      rq_wait_pos_spe_for_request(255, 204, 255, "1")
      rq_go_to("1")
      rq_wait("1")
      # end: URCap Program Node
      $ 2066 "Decap"
      $ 2067 "Action_Info≔'decapping'"
      global Action_Info="decapping"
      $ 2068 "Set GRP_3F_Enable=On"
      set_standard_digital_out(4, True)
      $ 2069 "Set GRP_3F_Decap=On"
      set_standard_digital_out(3, True)
      $ 2070 "Force"
      sleep(0.02)
      zero_ftsensor()
      force_mode(p[0.0,0.0,0.0,0.0,0.0,0.0], [0, 0, 1, 0, 0, 0], [0.0, 0.0, 1.0, 0.0, 0.0, 0.0], 2, [0.1, 0.1, 0.001, 0.3490658503988659, 0.3490658503988659, 0.3490658503988659])
      $ 2071 "check_decapping(offset=0.015, timeout=10, abort=CMD_Hold)" "noBreak"
      check_decapping(offset=0.015, timeout=10, abort=CMD_Hold)
      end_force_mode()
      stopl(5.0)
      $ 2072 "Set GRP_3F_Decap=Off"
      set_standard_digital_out(3, False)
      $ 2073 "Set GRP_3F_Enable=Off"
      set_standard_digital_out(4, False)
      $ 2074 "MoveL"
      $ 2075 "Waypoint_90" "breakAfter"
      movel(Waypoint_90_p, a=0.5, v=0.1, r=0.05)
      $ 2076 "MoveJ"
      $ 2077 "cap_dump_2" "breakAfter"
      movej(get_inverse_kin(cap_dump_2_p, qnear=cap_dump_2_q), a=0.5235987755982988, v=0.4363323129985824)
      # begin: URCap Program Node
      #   Source: Robotiq_Grippers, 3.17.0.105337, Robotiq Inc.
      #   Type: Gripper
      $ 2078 "Gripper Open (1)"
      if not(gripper_connected[0]):
        popup("Gripper 1 must be connected to run this program.", "No connection", False, True, True)
      end
      if not(rq_is_gripper_activated("1")):
        popup("Gripper 1 is not activated. Go to Installation tab > Gripper to activate it and run the program again.", "Not activated", False, True, True)
      end
      rq_set_pos_spd_for(0, 204, 255, "1")
      rq_wait_pos_spe_for_request(0, 204, 255, "1")
      rq_go_to("1")
      rq_wait("1")
      # end: URCap Program Node
      $ 2079 "MoveJ"
      $ 2080 "Waypoint_91" "breakAfter"
      movej(get_inverse_kin(Waypoint_91_p, qnear=Waypoint_91_q), a=0.5235987755982988, v=0.4363323129985824, r=0.036)
    elif (33 == switch_1):
      $ 2081 "Case 33"
      $ 2082 "Shake and liquid transfer"
      $ 2083 "MoveL"
      $ 2084 "Vial_liq_abov_1" "breakAfter"
      movel(Vial_liq_abov_1_p, a=0.5, v=0.1)
      $ 2085 "Vial_liq_pick_3" "breakAfter"
      movel(Vial_liq_pick_3_p, a=0.5, v=0.1)
      $ 2086 "Vial_liq_pick_4" "breakAfter"
      movel(Vial_liq_pick_4_p, a=0.5, v=0.1)
      # begin: URCap Program Node
      #   Source: Robotiq_Grippers, 3.17.0.105337, Robotiq Inc.
      #   Type: Gripper
      $ 2087 "Gripper Close (1)"
      if not(gripper_connected[0]):
        popup("Gripper 1 must be connected to run this program.", "No connection", False, True, True)
      end
      if not(rq_is_gripper_activated("1")):
        popup("Gripper 1 is not activated. Go to Installation tab > Gripper to activate it and run the program again.", "Not activated", False, True, True)
      end
      rq_set_pos_spd_for(255, 82, 71, "1")
      rq_wait_pos_spe_for_request(255, 82, 71, "1")
      rq_go_to("1")
      rq_wait("1")
      # end: URCap Program Node
      $ 2088 "Wait: 1.0"
      sleep(1.0)
      $ 2089 "Set GRP_3F_Open=On"
      set_standard_digital_out(5, True)
      $ 2090 "Wait: 0.5"
      sleep(0.5)
      $ 2091 "Vial_liq_abov_2" "breakAfter"
      movel(Vial_liq_abov_2_p, a=0.3, v=0.05, r=0.05)
      $ 2092 "MoveL"
      $ 2093 "Liquid_midway_1" "breakAfter"
      movel(Liquid_midway_1_p, a=0.5, v=0.1)
      $ 2094 "Loop 3 times"
      Loop_1 = 0
      while (Loop_1 < 3):
        $ 2095 "shake_3" "breakAfter"
        movel(shake_3_p, a=2.0, v=0.5)
        $ 2096 "shake_4" "breakAfter"
        movel(shake_4_p, a=2.0, v=0.5)
        Loop_1 = Loop_1 + 1
      end
      $ 2097 "drop_above_3" "breakAfter"
      movel(drop_above_3_p, a=0.5, v=0.1)
      $ 2098 "drop_above_4" "breakAfter"
      movel(drop_above_4_p, a=0.5, v=0.1)
      $ 2099 "liq_tran_3" "breakAfter"
      movel(liq_tran_3_p, a=0.5, v=0.05, r=0.008)
      $ 2100 "Wait: 1.0"
      sleep(1.0)
      $ 2101 "drop_above_5" "breakAfter"
      movel(drop_above_5_p, a=0.5, v=0.1)
      $ 2102 "Waypoint_92" "breakAfter"
      movel(Waypoint_92_p, a=0.5, v=0.1)
      $ 2103 "liq_tran_4" "breakAfter"
      movel(liq_tran_4_p, a=0.5, v=0.05)
      $ 2104 "Wait: 1.0"
      sleep(1.0)
      $ 2105 "drop_above_6" "breakAfter"
      movel(drop_above_6_p, a=0.5, v=0.1)
      $ 2106 "drop_above_7" "breakAfter"
      movel(drop_above_7_p, a=0.5, v=0.1)
      $ 2107 "Liquid_midway_2" "breakAfter"
      movel(Liquid_midway_2_p, a=0.5, v=0.1)
      $ 2108 "MoveL"
      $ 2109 "Vial_drop_abo_1" "breakAfter"
      movel(Vial_drop_abo_1_p, a=0.5, v=0.1)
      $ 2110 "Vial_liq_drop_1" "breakAfter"
      movel(Vial_liq_drop_1_p, a=0.5, v=0.1)
      # begin: URCap Program Node
      #   Source: Robotiq_Grippers, 3.17.0.105337, Robotiq Inc.
      #   Type: Gripper
      $ 2111 "Gripper Open (1)"
      if not(gripper_connected[0]):
        popup("Gripper 1 must be connected to run this program.", "No connection", False, True, True)
      end
      if not(rq_is_gripper_activated("1")):
        popup("Gripper 1 is not activated. Go to Installation tab > Gripper to activate it and run the program again.", "Not activated", False, True, True)
      end
      rq_set_pos_spd_for(0, 82, 71, "1")
      rq_wait_pos_spe_for_request(0, 82, 71, "1")
      rq_go_to("1")
      rq_wait("1")
      # end: URCap Program Node
      $ 2112 "Vial_drop_abo_2" "breakAfter"
      movel(Vial_drop_abo_2_p, a=0.5, v=0.1)
    elif (34 == switch_1):
      $ 2113 "Case 34"
      $ 2114 "Task≔'Dosing'"
      global Task="Dosing"
      $ 2115 "tilt_to_home()"
      tilt_to_home()
      $ 2116 "Powder dosing all"
      $ 2117 "tilt_angle_sent≔0.0"
      global tilt_angle_sent=0.0
      $ 2118 "send_target_info()"
      send_target_info()
      $ 2120 "prev_spat≔''"
      global prev_spat=""
      $ 2121 "spatula≔''"
      global spatula=""
      $ 2122 "scoop_status≔'normal'"
      global scoop_status="normal"
      $ 2123 "send_powder_info()"
      send_powder_info()
      $ 2124 "Set AO[0]=0.0"
      set_standard_analog_out(0, 0.0)
      $ 2125 "Wait: 0.2"
      sleep(0.2)
      $ 2126 "reach pots decapping pose"
      # begin: URCap Program Node
      #   Source: SensoPart VISOR Robotic, 2.0.6, SensoPart Industriesensorik GmbH
      #   Type: VISOR Robotic App
      $ 2132 "VISOR Easy Pick"
      def visorFuncEasyPick_e02a40():
        # begin: URCap Program Node
        #   Source: SensoPart VISOR Robotic, 2.0.6, SensoPart Industriesensorik GmbH
        #   Type: Easy Pick Setup
        $ 2133 "# 1 Setup" "noBreak"
        local easyPickVisorId = 1
        local easyPickArmMounted = True
        local easyPickSetJob = True
        local easyPickJobName = "Weight_scale"
        local easyPickAtImgAcq = False
        local easyPickImgAcqPose = Trigger
        # end: URCap Program Node
        # begin: URCap Program Node
        #   Source: SensoPart VISOR Robotic, 2.0.6, SensoPart Industriesensorik GmbH
        #   Type: Process
        $ 2134 "Process" "noBreak"
        local easyPickObjTaken = False
        local easyPickTrigger = False
        local easyPickPoseIdx = 0
        local easyPickPose = p[0,0,0,0,0,0]
        def easyPickFuncTrigger(visorId, setJob, jobName, arm):
        if (setJob):
          visor_changeJob(visorId, jobName, 6000)
        end
        if (arm):
          visor_trigger(visorId, 6000, "arm")
        else:
          visor_trigger(visorId, 6000)
        end
        global easyPickParts_4=visor_partsFound(visorId)
        visor_easyPickUpdate(visorId, "parts", visor_partsFound(visorId))
        return visor_getPose3d(visorId, 0)
      end
      while (not easyPickObjTaken):
        easyPickTrigger = (easyPickCount_4 >= visor_partsFound(easyPickVisorId)) or (easyPickCount_4 > 9) or (not visor_easyPickCheckIdent("02a34f", easyPickVisorId))
        if (easyPickTrigger):
          easyPickCount_4 = 0
        end
        easyPickPoseIdx = easyPickCount_4
        easyPickPose = visor_getPose3d(easyPickVisorId, easyPickPoseIdx)
        visor_easyPickUpdate(easyPickVisorId, "counter", easyPickPoseIdx)
        # begin: URCap Program Node
        #   Source: SensoPart VISOR Robotic, 2.0.6, SensoPart Industriesensorik GmbH
        #   Type: Image Acquisition Pose
        $ 2135 "Image Acquisition Pose" "noBreak"
        if (easyPickTrigger):
          if (not easyPickAtImgAcq):
            movej(pose_trans(easyPickImgAcqPose,p[0.0000,0.0000,-0.0000,0.0000,0.0000,0.0000]),a=1.3963,v=1.0472,t=0.000000,r=0.000000)
            easyPickAtImgAcq = True
          end
          easyPickPose = easyPickFuncTrigger(easyPickVisorId, easyPickSetJob, easyPickJobName, easyPickArmMounted)
        end
        # end: URCap Program Node
        # begin: URCap Program Node
        #   Source: SensoPart VISOR Robotic, 2.0.6, SensoPart Industriesensorik GmbH
        #   Type: Object Detected
        $ 2136 "Object Detected" "noBreak"
        if (visor_partsFound(easyPickVisorId) > 0):
          $ 2137 "Open Gripper" "noBreak"
          $ 2138 "weight_value≔get_weight()" "noBreak"
          global weight_value=get_weight()
          $ 2139 "Wait: 0.5" "noBreak"
          sleep(0.5)
          $ 2140 "diff≔target_weight-weight_value" "noBreak"
          global diff=target_weight-weight_value
          $ 2141 "compute_level_percent(W_now, weight_value)" "noBreak"
          compute_level_percent(W_now, weight_value)
          $ 2142 "send_level_info()" "noBreak"
          send_level_info()
          $ 2143 "spatula≔select_spatula(Flowability, level, diff, bulk_density, mouth_d)" "noBreak"
          global spatula=select_spatula(Flowability, level, diff, bulk_density, mouth_d)
          $ 2144 "Wait: 0.2" "noBreak"
          sleep(0.2)
          $ 2145 "send_spatula_info()" "noBreak"
          send_spatula_info()
          $ 2146 "Pick spatula" "noBreak"
          $ 2147 "If spatula ≟ 'spatula_L'" "noBreak"
          if (spatula  ==  "spatula_L"):
            $ 2148 "MoveJ" "noBreak"
            $ 2149 "Spatula_otw" "noBreak"
            movej(get_inverse_kin(Spatula_otw_p, qnear=Spatula_otw_q), a=1.3962634015954636, v=1.0471975511965976)
            $ 2150 "pick_spat_L_abv" "noBreak"
            movej(get_inverse_kin(pick_spat_L_abv_p, qnear=pick_spat_L_abv_q), a=1.3962634015954636, v=1.0471975511965976)
            $ 2151 "MoveL" "noBreak"
            $ 2152 "spat_L_pick" "noBreak"
            movel(spat_L_pick_p, a=1.2, v=0.25)
            # begin: URCap Program Node
            #   Source: Robotiq_Grippers, 3.17.0.105337, Robotiq Inc.
            #   Type: Gripper
            $ 2153 "Gripper Close (1)" "noBreak"
            if not(gripper_connected[0]):
              popup("Gripper 1 must be connected to run this program.", "No connection", False, True, True)
            end
            if not(rq_is_gripper_activated("1")):
              popup("Gripper 1 is not activated. Go to Installation tab > Gripper to activate it and run the program again.", "Not activated", False, True, True)
            end
            rq_set_pos_spd_for(255, 0, 77, "1")
            rq_wait_pos_spe_for_request(255, 0, 77, "1")
            rq_go_to("1")
            rq_wait("1")
            # end: URCap Program Node
            $ 2154 "spat_L_lift" "noBreak"
            movel(spat_L_lift_p, a=1.2, v=0.25, r=0.01)
            $ 2155 "spat_L_side" "noBreak"
            movel(spat_L_side_p, a=1.2, v=0.25, r=0.01)
            $ 2156 "spat_L_up" "noBreak"
            movel(spat_L_up_p, a=1.2, v=0.25, r=0.05)
            $ 2157 "MoveJ" "noBreak"
            $ 2158 "Spatula_otw" "noBreak"
            movej(get_inverse_kin(Spatula_otw_p, qnear=Spatula_otw_q), a=1.3962634015954636, v=1.0471975511965976)
          else:
            $ 2159 "ElseIf spatula ≟'spatula_M'" "noBreak"
            if (spatula  == "spatula_M"):
              $ 2160 "MoveJ" "noBreak"
              $ 2161 "Spatula_otw" "noBreak"
              movej(get_inverse_kin(Spatula_otw_p, qnear=Spatula_otw_q), a=1.3962634015954636, v=1.0471975511965976)
              $ 2162 "spat_M_up" "noBreak"
              movej(get_inverse_kin(spat_M_up_p, qnear=spat_M_up_q), a=1.3962634015954636, v=1.0471975511965976, r=0.05)
              $ 2163 "MoveL" "noBreak"
              $ 2164 "spat_M_pick" "noBreak"
              movel(spat_M_pick_p, a=1.2, v=0.25)
              # begin: URCap Program Node
              #   Source: Robotiq_Grippers, 3.17.0.105337, Robotiq Inc.
              #   Type: Gripper
              $ 2165 "Gripper Close (1)" "noBreak"
              if not(gripper_connected[0]):
                popup("Gripper 1 must be connected to run this program.", "No connection", False, True, True)
              end
              if not(rq_is_gripper_activated("1")):
                popup("Gripper 1 is not activated. Go to Installation tab > Gripper to activate it and run the program again.", "Not activated", False, True, True)
              end
              rq_set_pos_spd_for(255, 0, 77, "1")
              rq_wait_pos_spe_for_request(255, 0, 77, "1")
              rq_go_to("1")
              rq_wait("1")
              # end: URCap Program Node
              $ 2166 "spat_M_up" "noBreak"
              movel(spat_M_up_p, a=1.2, v=0.25, r=0.05)
              $ 2167 "Spatula_otw" "noBreak"
              movel(Spatula_otw_p, a=1.2, v=0.25)
              $ 2168 "switch_spat_M≔ False " "noBreak"
              global switch_spat_M=  False
            else:
              $ 2169 "ElseIf spatula≟'spatula_S'" "noBreak"
              if (spatula == "spatula_S"):
                $ 2170 "MoveJ" "noBreak"
                $ 2171 "Spatula_otw" "noBreak"
                movej(get_inverse_kin(Spatula_otw_p, qnear=Spatula_otw_q), a=1.3962634015954636, v=1.0471975511965976)
                $ 2172 "spat_S_Up_7" "noBreak"
                movej(get_inverse_kin(spat_S_Up_7_p, qnear=spat_S_Up_7_q), a=1.3962634015954636, v=1.0471975511965976, r=0.05)
                $ 2173 "MoveL" "noBreak"
                $ 2174 "spat_S_Pick_4" "noBreak"
                movel(spat_S_Pick_4_p, a=1.2, v=0.25)
                # begin: URCap Program Node
                #   Source: Robotiq_Grippers, 3.17.0.105337, Robotiq Inc.
                #   Type: Gripper
                $ 2175 "Gripper Close (1)" "noBreak"
                if not(gripper_connected[0]):
                  popup("Gripper 1 must be connected to run this program.", "No connection", False, True, True)
                end
                if not(rq_is_gripper_activated("1")):
                  popup("Gripper 1 is not activated. Go to Installation tab > Gripper to activate it and run the program again.", "Not activated", False, True, True)
                end
                rq_set_pos_spd_for(255, 0, 77, "1")
                rq_wait_pos_spe_for_request(255, 0, 77, "1")
                rq_go_to("1")
                rq_wait("1")
                # end: URCap Program Node
                $ 2176 "spat_S_Up_8" "noBreak"
                movel(spat_S_Up_8_p, a=1.2, v=0.25, r=0.05)
                $ 2177 "Spatula_otw" "noBreak"
                movel(Spatula_otw_p, a=1.2, v=0.25)
                $ 2178 "switch_spat_S≔ False " "noBreak"
                global switch_spat_S=  False
              else:
                $ 2179 "ElseIf spatula≟'spatula_flat_M'" "noBreak"
                if (spatula == "spatula_flat_M"):
                  $ 2180 "MoveJ" "noBreak"
                  $ 2181 "Spatula_otw" "noBreak"
                  movej(get_inverse_kin(Spatula_otw_p, qnear=Spatula_otw_q), a=1.3962634015954636, v=1.0471975511965976)
                  $ 2182 "spat_flatM_up" "noBreak"
                  movej(get_inverse_kin(spat_flatM_up_p, qnear=spat_flatM_up_q), a=1.3962634015954636, v=1.0471975511965976, r=0.05)
                  $ 2183 "MoveL" "noBreak"
                  $ 2184 "spat_flatM_pick" "noBreak"
                  movel(spat_flatM_pick_p, a=1.2, v=0.25)
                  # begin: URCap Program Node
                  #   Source: Robotiq_Grippers, 3.17.0.105337, Robotiq Inc.
                  #   Type: Gripper
                  $ 2185 "Gripper Close (1)" "noBreak"
                  if not(gripper_connected[0]):
                    popup("Gripper 1 must be connected to run this program.", "No connection", False, True, True)
                  end
                  if not(rq_is_gripper_activated("1")):
                    popup("Gripper 1 is not activated. Go to Installation tab > Gripper to activate it and run the program again.", "Not activated", False, True, True)
                  end
                  rq_set_pos_spd_for(255, 0, 77, "1")
                  rq_wait_pos_spe_for_request(255, 0, 77, "1")
                  rq_go_to("1")
                  rq_wait("1")
                  # end: URCap Program Node
                  $ 2186 "spat_flatM_up" "noBreak"
                  movel(spat_flatM_up_p, a=1.2, v=0.25, r=0.05)
                  $ 2187 "Spatula_otw" "noBreak"
                  movel(Spatula_otw_p, a=1.2, v=0.25)
                  $ 2188 "switch_spat_F_M≔ False " "noBreak"
                  global switch_spat_F_M=  False
                else:
                  $ 2189 "ElseIf spatula≟'spatula_flat_S'" "noBreak"
                  if (spatula == "spatula_flat_S"):
                    $ 2190 "MoveJ" "noBreak"
                    $ 2191 "Spatula_otw" "noBreak"
                    movej(get_inverse_kin(Spatula_otw_p, qnear=Spatula_otw_q), a=1.3962634015954636, v=1.0471975511965976)
                    $ 2192 "spat_flatS_up" "noBreak"
                    movej(get_inverse_kin(spat_flatS_up_p, qnear=spat_flatS_up_q), a=1.3962634015954636, v=1.0471975511965976, r=0.05)
                    $ 2193 "MoveL" "noBreak"
                    $ 2194 "spat_flatS_pick" "noBreak"
                    movel(spat_flatS_pick_p, a=1.2, v=0.25)
                    # begin: URCap Program Node
                    #   Source: Robotiq_Grippers, 3.17.0.105337, Robotiq Inc.
                    #   Type: Gripper
                    $ 2195 "Gripper Close (1)" "noBreak"
                    if not(gripper_connected[0]):
                      popup("Gripper 1 must be connected to run this program.", "No connection", False, True, True)
                    end
                    if not(rq_is_gripper_activated("1")):
                      popup("Gripper 1 is not activated. Go to Installation tab > Gripper to activate it and run the program again.", "Not activated", False, True, True)
                    end
                    rq_set_pos_spd_for(255, 0, 77, "1")
                    rq_wait_pos_spe_for_request(255, 0, 77, "1")
                    rq_go_to("1")
                    rq_wait("1")
                    # end: URCap Program Node
                    $ 2196 "spat_flatS_up" "noBreak"
                    movel(spat_flatS_up_p, a=1.2, v=0.25, r=0.05)
                    $ 2197 "Spatula_otw" "noBreak"
                    movel(Spatula_otw_p, a=1.2, v=0.25)
                    $ 2198 "switch_spat_F_S≔ False " "noBreak"
                    global switch_spat_F_S=  False
                  end
                end
              end
            end
          end
          $ 2199 "Action_Info≔'Scooping'" "noBreak"
          global Action_Info="Scooping"
          $ 2200 "auto_tilt_and_scoop(W_now, target_weight, weight_value)" "noBreak"
          auto_tilt_and_scoop(W_now, target_weight, weight_value)
          $ 2201 "Action_Info≔'Dosing'" "noBreak"
          global Action_Info="Dosing"
          # begin: URCap Program Node
          #   Source: SensoPart VISOR Robotic, 2.0.6, SensoPart Industriesensorik GmbH
          #   Type: Approach Pose
          $ 2202 "Approach Pose" "noBreak"
          movej(pose_trans(easyPickPose,p[0.0000,0.0000,-0.0000,0.0000,0.0000,0.0000]),a=0.2618,v=0.1745,t=0.000000,r=0.000000)
          # end: URCap Program Node
          # begin: URCap Program Node
          #   Source: SensoPart VISOR Robotic, 2.0.6, SensoPart Industriesensorik GmbH
          #   Type: Target Pose
          $ 2203 "Target Pose" "noBreak"
          movel(pose_trans(easyPickPose,p[0.0000,0.0000,-0.0000,0.0000,0.0000,0.0000]),a=0.0500,v=0.0200,t=0.000000,r=0.000000)
          # end: URCap Program Node
          $ 2204 "Close Gripper" "noBreak"
          $ 2205 "current_p≔get_actual_tcp_pose()" "noBreak"
          global current_p= get_actual_tcp_pose ()
          $ 2206 "dispense_pos≔pose_trans(current_p,p[0,0,0,0,-deg2rad(spatula_ry),0])" "noBreak"
          global dispense_pos=pose_trans(current_p,p[0,0,0,0,-deg2rad(spatula_ry),0])
          $ 2207 "Loop weight_value≤target_weight and delta_count≤3" "noBreak"
          thread Thread_while_2207():
            while (True):
              $ 2208 "MoveL" "noBreak"
              $ 2209 "dispense_pos" "noBreak"
              movel(dispense_pos, a=0.2, v=0.1)
              $ 2210 "log_weight()" "noBreak"
              log_weight()
              $ 2212 "CCW_full_Rotate()" "noBreak"
              CCW_full_Rotate()
              $ 2213 "Start_thread≔ True " "noBreak"
              global Start_thread=  True
              $ 2214 "vib_thread≔ True " "noBreak"
              global vib_thread=  True
              $ 2215 "Wait: 0.5" "noBreak"
              sleep(0.5)
              $ 2216 "If diff ≥(target_g*1.2)" "noBreak"
              if (diff  >= (target_g*1.2)):
                $ 2217 "tilt_pose≔pose_trans(get_actual_tcp_pose(), p[0, 0, 0, 0, 0, 2.0])" "noBreak"
                global tilt_pose=pose_trans(get_actual_tcp_pose(), p[0, 0, 0, 0, 0, 2.0])
                $ 2218 "movel(tilt_pose, a=0.5, v=0.5, r=0.00001)" "noBreak"
                movel(tilt_pose, a=0.5, v=0.5, r=0.00001)
              else:
                $ 2219 "Else" "noBreak"
                $ 2220 "Loop weight_value≤(target_weight-0.00) and tilt_angle≥(-1.999) and tilt_angle≤0.5" "noBreak"
                thread Thread_while_2220():
                  while (True):
                    $ 2221 "current_error≔target_weight-weight_value" "noBreak"
                    global current_error=target_weight-weight_value
                    $ 2222 "Integral_error≔Integral_error+current_error*dt" "noBreak"
                    global Integral_error=Integral_error+current_error*dt
                    $ 2223 "derivative≔(current_error-previous_error)/dt" "noBreak"
                    global derivative=(current_error-previous_error)/dt
                    $ 2224 "tilt_increment≔(kp*current_error)+(ki*Integral_error)+(kd*derivative)" "noBreak"
                    global tilt_increment=(kp*current_error)+(ki*Integral_error)+(kd*derivative)
                    $ 2225 "current_pose≔get_actual_tcp_pose()" "noBreak"
                    global current_pose= get_actual_tcp_pose ()
                    $ 2226 "tilt_angle≔current_pose[5]" "noBreak"
                    global tilt_angle=current_pose[5]
                    $ 2227 "tilt_pose≔pose_trans(current_pose, p[0, 0, 0, 0, 0, tilt_increment])" "noBreak"
                    global tilt_pose=pose_trans(current_pose, p[0, 0, 0, 0, 0, tilt_increment])
                    $ 2228 "movel(tilt_pose, a=0.1, v=0.1, r=0.00001)" "noBreak"
                    movel(tilt_pose, a=0.1, v=0.1, r=0.00001)
                    $ 2229 "previous_error≔current_error" "noBreak"
                    global previous_error=current_error
                  end
                end
                if (weight_value <= (target_weight-0.00)  and  tilt_angle >= (-1.999)  and  tilt_angle <= 0.5):
                  global thread_handler_2220=run Thread_while_2220()
                  while (weight_value <= (target_weight-0.00)  and  tilt_angle >= (-1.999)  and  tilt_angle <= 0.5):
                    sync()
                  end
                  kill thread_handler_2220
                end
              end
              $ 2230 "weight_value≔get_weight()" "noBreak"
              global weight_value=get_weight()
              $ 2231 "tilt_angle≔-1" "noBreak"
              global tilt_angle=-1
              $ 2232 "Wait: 0.5" "noBreak"
              sleep(0.5)
              $ 2233 "Start_thread≔ False " "noBreak"
              global Start_thread=  False
              $ 2234 "vib_thread≔ False " "noBreak"
              global vib_thread=  False
              $ 2235 "dispense_pos" "noBreak"
              movel(dispense_pos, a=1.2, v=0.25)
              $ 2236 "compute_level_percent(W_now, weight_value)" "noBreak"
              compute_level_percent(W_now, weight_value)
              $ 2237 "If delta<0.01" "noBreak"
              if (delta<0.01):
                $ 2238 "delta_count≔delta_count+1" "noBreak"
                global delta_count=delta_count+1
              else:
                $ 2239 "Else" "noBreak"
                $ 2240 "delta_count≔0" "noBreak"
                global delta_count=0
              end
              $ 2241 "prev_spat≔spatula" "noBreak"
              global prev_spat=spatula
              $ 2242 "Wait: 0.2" "noBreak"
              sleep(0.2)
              $ 2243 "spatula≔select_spatula(Flowability, level, diff, bulk_density, mouth_d)" "noBreak"
              global spatula=select_spatula(Flowability, level, diff, bulk_density, mouth_d)
              $ 2244 "Wait: 1.0" "noBreak"
              sleep(1.0)
              $ 2245 "send_level_info()" "noBreak"
              send_level_info()
              $ 2246 "send_spatula_info()" "noBreak"
              send_spatula_info()
              $ 2247 "Integral_error≔0" "noBreak"
              global Integral_error=0
              $ 2248 "current_error≔0" "noBreak"
              global current_error=0
              $ 2249 "previous_error≔0" "noBreak"
              global previous_error=0
              $ 2250 "Set AO[0]=0.0" "noBreak"
              set_standard_analog_out(0, 0.0)
              $ 2251 "Wait: 0.5" "noBreak"
              sleep(0.5)
              $ 2252 "swtich spatula" "noBreak"
              $ 2253 "If spatula ≟ 'spatula_M' and switch_spat_M≟ True " "noBreak"
              if (spatula  ==  "spatula_M"  and  switch_spat_M ==   True  ):
                $ 2254 "MoveJ" "noBreak"
                $ 2255 "Spatula_otw" "noBreak"
                movej(get_inverse_kin(Spatula_otw_p, qnear=Spatula_otw_q), a=1.3962634015954636, v=1.0471975511965976)
                $ 2256 "spat_L_up" "noBreak"
                movej(get_inverse_kin(spat_L_up_p, qnear=spat_L_up_q), a=1.3962634015954636, v=1.0471975511965976)
                $ 2257 "MoveL" "noBreak"
                $ 2258 "spat_L_side" "noBreak"
                movel(spat_L_side_p, a=1.2, v=0.25)
                $ 2259 "spat_L_lift" "noBreak"
                movel(spat_L_lift_p, a=1.2, v=0.25)
                $ 2260 "spat_L_pick" "noBreak"
                movel(spat_L_pick_p, a=0.2, v=0.1)
                # begin: URCap Program Node
                #   Source: Robotiq_Grippers, 3.17.0.105337, Robotiq Inc.
                #   Type: Gripper
                $ 2261 "Gripper Open (1)" "noBreak"
                if not(gripper_connected[0]):
                  popup("Gripper 1 must be connected to run this program.", "No connection", False, True, True)
                end
                if not(rq_is_gripper_activated("1")):
                  popup("Gripper 1 is not activated. Go to Installation tab > Gripper to activate it and run the program again.", "Not activated", False, True, True)
                end
                rq_set_pos_spd_for(0, 255, 77, "1")
                rq_wait_pos_spe_for_request(0, 255, 77, "1")
                rq_go_to("1")
                rq_wait("1")
                # end: URCap Program Node
                $ 2262 "spat_M_pick" "noBreak"
                movel(spat_M_pick_p, a=1.2, v=0.25)
                # begin: URCap Program Node
                #   Source: Robotiq_Grippers, 3.17.0.105337, Robotiq Inc.
                #   Type: Gripper
                $ 2263 "Gripper Close (1)" "noBreak"
                if not(gripper_connected[0]):
                  popup("Gripper 1 must be connected to run this program.", "No connection", False, True, True)
                end
                if not(rq_is_gripper_activated("1")):
                  popup("Gripper 1 is not activated. Go to Installation tab > Gripper to activate it and run the program again.", "Not activated", False, True, True)
                end
                rq_set_pos_spd_for(255, 0, 77, "1")
                rq_wait_pos_spe_for_request(255, 0, 77, "1")
                rq_go_to("1")
                rq_wait("1")
                # end: URCap Program Node
                $ 2264 "spat_M_up" "noBreak"
                movel(spat_M_up_p, a=1.2, v=0.25)
                $ 2265 "Spatula_otw" "noBreak"
                movel(Spatula_otw_p, a=1.2, v=0.25)
                $ 2266 "switch_spat_M≔ False " "noBreak"
                global switch_spat_M=  False
                $ 2267 "correction_reset()" "noBreak"
                correction_reset()
              else:
                $ 2268 "ElseIf spatula ≟ 'spatula_S' and switch_spat_S ≟ True and prev_spat≟'spatula_M'" "noBreak"
                if (spatula  ==  "spatula_S" and switch_spat_S  ==   True  and prev_spat == "spatula_M"):
                  $ 2269 "MoveL" "noBreak"
                  $ 2270 "Spatula_otw" "noBreak"
                  movel(Spatula_otw_p, a=1.2, v=0.25)
                  $ 2271 "spat_M_up" "noBreak"
                  movel(spat_M_up_p, a=1.2, v=0.25)
                  $ 2272 "spat_M_pick" "noBreak"
                  movel(spat_M_pick_p, a=0.2, v=0.1)
                  # begin: URCap Program Node
                  #   Source: Robotiq_Grippers, 3.17.0.105337, Robotiq Inc.
                  #   Type: Gripper
                  $ 2273 "Gripper Open (1)" "noBreak"
                  if not(gripper_connected[0]):
                    popup("Gripper 1 must be connected to run this program.", "No connection", False, True, True)
                  end
                  if not(rq_is_gripper_activated("1")):
                    popup("Gripper 1 is not activated. Go to Installation tab > Gripper to activate it and run the program again.", "Not activated", False, True, True)
                  end
                  rq_set_pos_spd_for(0, 255, 77, "1")
                  rq_wait_pos_spe_for_request(0, 255, 77, "1")
                  rq_go_to("1")
                  rq_wait("1")
                  # end: URCap Program Node
                  $ 2274 "spat_S_pick" "noBreak"
                  movel(spat_S_pick_p, a=1.2, v=0.25)
                  # begin: URCap Program Node
                  #   Source: Robotiq_Grippers, 3.17.0.105337, Robotiq Inc.
                  #   Type: Gripper
                  $ 2275 "Gripper Close (1)" "noBreak"
                  if not(gripper_connected[0]):
                    popup("Gripper 1 must be connected to run this program.", "No connection", False, True, True)
                  end
                  if not(rq_is_gripper_activated("1")):
                    popup("Gripper 1 is not activated. Go to Installation tab > Gripper to activate it and run the program again.", "Not activated", False, True, True)
                  end
                  rq_set_pos_spd_for(255, 0, 77, "1")
                  rq_wait_pos_spe_for_request(255, 0, 77, "1")
                  rq_go_to("1")
                  rq_wait("1")
                  # end: URCap Program Node
                  $ 2276 "spat_S_up" "noBreak"
                  movel(spat_S_up_p, a=1.2, v=0.25)
                  $ 2277 "Spatula_otw" "noBreak"
                  movel(Spatula_otw_p, a=1.2, v=0.25)
                  $ 2278 "switch_spat_S≔ False " "noBreak"
                  global switch_spat_S=  False
                  $ 2279 "correction_reset()" "noBreak"
                  correction_reset()
                else:
                  $ 2280 "ElseIf spatula≟'spatula_S' and switch_spat_S≟ True  and prev_spat≟'spatula_L'" "noBreak"
                  if (spatula == "spatula_S" and switch_spat_S ==   True    and  prev_spat == "spatula_L"):
                    $ 2281 "MoveJ" "noBreak"
                    $ 2282 "Spatula_otw" "noBreak"
                    movej(get_inverse_kin(Spatula_otw_p, qnear=Spatula_otw_q), a=1.3962634015954636, v=1.0471975511965976)
                    $ 2283 "spat_L_up" "noBreak"
                    movej(get_inverse_kin(spat_L_up_p, qnear=spat_L_up_q), a=1.3962634015954636, v=1.0471975511965976)
                    $ 2284 "MoveL" "noBreak"
                    $ 2285 "spat_L_side" "noBreak"
                    movel(spat_L_side_p, a=1.2, v=0.25)
                    $ 2286 "spat_L_lift" "noBreak"
                    movel(spat_L_lift_p, a=1.2, v=0.25)
                    $ 2287 "spat_L_pick" "noBreak"
                    movel(spat_L_pick_p, a=0.2, v=0.1)
                    # begin: URCap Program Node
                    #   Source: Robotiq_Grippers, 3.17.0.105337, Robotiq Inc.
                    #   Type: Gripper
                    $ 2288 "Gripper Open (1)" "noBreak"
                    if not(gripper_connected[0]):
                      popup("Gripper 1 must be connected to run this program.", "No connection", False, True, True)
                    end
                    if not(rq_is_gripper_activated("1")):
                      popup("Gripper 1 is not activated. Go to Installation tab > Gripper to activate it and run the program again.", "Not activated", False, True, True)
                    end
                    rq_set_pos_spd_for(0, 255, 77, "1")
                    rq_wait_pos_spe_for_request(0, 255, 77, "1")
                    rq_go_to("1")
                    rq_wait("1")
                    # end: URCap Program Node
                    $ 2289 "spat_S_pick" "noBreak"
                    movel(spat_S_pick_p, a=1.2, v=0.25)
                    # begin: URCap Program Node
                    #   Source: Robotiq_Grippers, 3.17.0.105337, Robotiq Inc.
                    #   Type: Gripper
                    $ 2290 "Gripper Close (1)" "noBreak"
                    if not(gripper_connected[0]):
                      popup("Gripper 1 must be connected to run this program.", "No connection", False, True, True)
                    end
                    if not(rq_is_gripper_activated("1")):
                      popup("Gripper 1 is not activated. Go to Installation tab > Gripper to activate it and run the program again.", "Not activated", False, True, True)
                    end
                    rq_set_pos_spd_for(255, 0, 77, "1")
                    rq_wait_pos_spe_for_request(255, 0, 77, "1")
                    rq_go_to("1")
                    rq_wait("1")
                    # end: URCap Program Node
                    $ 2291 "spat_S_up" "noBreak"
                    movel(spat_S_up_p, a=1.2, v=0.25)
                    $ 2292 "Spatula_otw" "noBreak"
                    movel(Spatula_otw_p, a=1.2, v=0.25)
                    $ 2293 "switch_spat_S≔ False " "noBreak"
                    global switch_spat_S=  False
                    $ 2294 "correction_reset()" "noBreak"
                    correction_reset()
                  else:
                    $ 2295 "ElseIf spatula≟'spatula_flat_S'  and switch_spat_F_S ≟ True " "noBreak"
                    if (spatula == "spatula_flat_S"   and  switch_spat_F_S  ==   True  ):
                      $ 2296 "MoveL" "noBreak"
                      $ 2297 "Spatula_otw" "noBreak"
                      movel(Spatula_otw_p, a=1.2, v=0.25)
                      $ 2298 "spat_flatM_up" "noBreak"
                      movel(spat_flatM_up_p, a=1.2, v=0.25)
                      $ 2299 "spat_flatM_pick" "noBreak"
                      movel(spat_flatM_pick_p, a=0.2, v=0.1)
                      # begin: URCap Program Node
                      #   Source: Robotiq_Grippers, 3.17.0.105337, Robotiq Inc.
                      #   Type: Gripper
                      $ 2300 "Gripper Open (1)" "noBreak"
                      if not(gripper_connected[0]):
                        popup("Gripper 1 must be connected to run this program.", "No connection", False, True, True)
                      end
                      if not(rq_is_gripper_activated("1")):
                        popup("Gripper 1 is not activated. Go to Installation tab > Gripper to activate it and run the program again.", "Not activated", False, True, True)
                      end
                      rq_set_pos_spd_for(0, 255, 74, "1")
                      rq_wait_pos_spe_for_request(0, 255, 74, "1")
                      rq_go_to("1")
                      rq_wait("1")
                      # end: URCap Program Node
                      $ 2301 "spat_flatS_pick" "noBreak"
                      movel(spat_flatS_pick_p, a=1.2, v=0.25)
                      # begin: URCap Program Node
                      #   Source: Robotiq_Grippers, 3.17.0.105337, Robotiq Inc.
                      #   Type: Gripper
                      $ 2302 "Gripper Close (1)" "noBreak"
                      if not(gripper_connected[0]):
                        popup("Gripper 1 must be connected to run this program.", "No connection", False, True, True)
                      end
                      if not(rq_is_gripper_activated("1")):
                        popup("Gripper 1 is not activated. Go to Installation tab > Gripper to activate it and run the program again.", "Not activated", False, True, True)
                      end
                      rq_set_pos_spd_for(255, 0, 77, "1")
                      rq_wait_pos_spe_for_request(255, 0, 77, "1")
                      rq_go_to("1")
                      rq_wait("1")
                      # end: URCap Program Node
                      $ 2303 "spat_flatS_up" "noBreak"
                      movel(spat_flatS_up_p, a=1.2, v=0.25)
                      $ 2304 "Spatula_otw" "noBreak"
                      movel(Spatula_otw_p, a=1.2, v=0.25)
                      $ 2305 "switch_spat_F_S≔ False " "noBreak"
                      global switch_spat_F_S=  False
                      $ 2306 "correction_reset()" "noBreak"
                      correction_reset()
                    end
                  end
                end
              end
              $ 2307 "tilt(level)" "noBreak"
              tilt(level)
              $ 2308 "Action_Info≔'Scooping'" "noBreak"
              global Action_Info="Scooping"
              $ 2309 "auto_tilt_and_scoop(W_now, target_weight, weight_value)" "noBreak"
              auto_tilt_and_scoop(W_now, target_weight, weight_value)
              $ 2310 "Action_Info≔'Dosing'" "noBreak"
              global Action_Info="Dosing"
            end
          end
          if (weight_value <= target_weight and delta_count <= 3):
            global thread_handler_2207=run Thread_while_2207()
            while (weight_value <= target_weight and delta_count <= 3):
              sync()
            end
            kill thread_handler_2207
          end
          $ 2311 "Start_thread≔ False " "noBreak"
          global Start_thread=  False
          $ 2312 "vib_thread≔ False " "noBreak"
          global vib_thread=  False
          # begin: URCap Program Node
          #   Source: SensoPart VISOR Robotic, 2.0.6, SensoPart Industriesensorik GmbH
          #   Type: Exit Pose
          $ 2313 "Exit Pose" "noBreak"
          movel(pose_trans(easyPickPose,p[0.0000,0.0000,-0.0000,0.0000,0.0000,0.0000]),a=0.5000,v=0.2500,t=0.000000,r=0.000000)
          # end: URCap Program Node
          easyPickObjTaken = True
        end
        # end: URCap Program Node
        # begin: URCap Program Node
        #   Source: SensoPart VISOR Robotic, 2.0.6, SensoPart Industriesensorik GmbH
        #   Type: No Object Detected
        $ 2314 "No Object Detected" "noBreak"
        if (visor_partsFound(easyPickVisorId) < 1):
          $ 2315 "Popup: No weigh scale detected" "noBreak"
          popup("No weigh scale detected", "Message", False, False, blocking=True)
          else:
        end
        # end: URCap Program Node
      end
      easyPickCount_4 = easyPickCount_4 + 1
      visor_easyPickUpdate(easyPickVisorId, "counter", easyPickCount_4)
      visor_easyPickSetIdent("02a34f", easyPickVisorId)
      # end: URCap Program Node
    end
    visorFuncEasyPick_e02a40()
    # end: URCap Program Node
    $ 2316 "MoveL"
    $ 2317 "dispense_pos" "breakAfter"
    movel(dispense_pos, a=0.2, v=0.1)
    $ 2318 "after_scoop()"
    after_scoop()
    $ 2319 "Place spatula back to the rack"
    $ 2320 "If spatula ≟ 'spatula_L'"
    if (spatula  ==  "spatula_L"):
      $ 2321 "MoveJ"
      $ 2322 "Spatula_otw" "breakAfter"
      movej(get_inverse_kin(Spatula_otw_p, qnear=Spatula_otw_q), a=1.3962634015954636, v=1.0471975511965976)
      $ 2323 "MoveL"
      $ 2324 "spat_L_up" "breakAfter"
      movel(spat_L_up_p, a=1.2, v=0.25, r=0.05)
      $ 2325 "spat_L_side" "breakAfter"
      movel(spat_L_side_p, a=1.2, v=0.25, r=0.01)
      $ 2326 "spat_L_lift" "breakAfter"
      movel(spat_L_lift_p, a=1.2, v=0.25, r=0.01)
      $ 2327 "spat_L_pick" "breakAfter"
      movel(spat_L_pick_p, a=0.2, v=0.1)
      # begin: URCap Program Node
      #   Source: Robotiq_Grippers, 3.17.0.105337, Robotiq Inc.
      #   Type: Gripper
      $ 2328 "Gripper Open (1)"
      if not(gripper_connected[0]):
        popup("Gripper 1 must be connected to run this program.", "No connection", False, True, True)
      end
      if not(rq_is_gripper_activated("1")):
        popup("Gripper 1 is not activated. Go to Installation tab > Gripper to activate it and run the program again.", "Not activated", False, True, True)
      end
      rq_set_pos_spd_for(0, 128, 128, "1")
      rq_wait_pos_spe_for_request(0, 128, 128, "1")
      rq_go_to("1")
      rq_wait("1")
      # end: URCap Program Node
      $ 2329 "MoveJ"
      $ 2330 "pick_spat_L_abv" "breakAfter"
      movej(get_inverse_kin(pick_spat_L_abv_p, qnear=pick_spat_L_abv_q), a=1.3962634015954636, v=1.0471975511965976)
      $ 2331 "Spatula_otw" "breakAfter"
      movej(get_inverse_kin(Spatula_otw_p, qnear=Spatula_otw_q), a=1.3962634015954636, v=1.0471975511965976)
    else:
      $ 2332 "ElseIf spatula ≟'spatula_M'"
      if (spatula  == "spatula_M"):
        $ 2333 "MoveJ"
        $ 2334 "Spatula_otw" "breakAfter"
        movej(get_inverse_kin(Spatula_otw_p, qnear=Spatula_otw_q), a=1.3962634015954636, v=1.0471975511965976)
        $ 2335 "spat_M_up" "breakAfter"
        movej(get_inverse_kin(spat_M_up_p, qnear=spat_M_up_q), a=1.3962634015954636, v=1.0471975511965976, r=0.05)
        $ 2336 "MoveL"
        $ 2337 "spat_M_pick" "breakAfter"
        movel(spat_M_pick_p, a=0.2, v=0.1)
        # begin: URCap Program Node
        #   Source: Robotiq_Grippers, 3.17.0.105337, Robotiq Inc.
        #   Type: Gripper
        $ 2338 "Gripper Open (1)"
        if not(gripper_connected[0]):
          popup("Gripper 1 must be connected to run this program.", "No connection", False, True, True)
        end
        if not(rq_is_gripper_activated("1")):
          popup("Gripper 1 is not activated. Go to Installation tab > Gripper to activate it and run the program again.", "Not activated", False, True, True)
        end
        rq_set_pos_spd_for(0, 128, 128, "1")
        rq_wait_pos_spe_for_request(0, 128, 128, "1")
        rq_go_to("1")
        rq_wait("1")
        # end: URCap Program Node
        $ 2339 "spat_M_up" "breakAfter"
        movel(spat_M_up_p, a=1.2, v=0.25, r=0.05)
        $ 2340 "Spatula_otw" "breakAfter"
        movel(Spatula_otw_p, a=1.2, v=0.25)
        $ 2341 "switch_spat_M≔ False "
        global switch_spat_M=  False
      else:
        $ 2342 "ElseIf spatula≟'spatula_S'"
        if (spatula == "spatula_S"):
          $ 2343 "MoveJ"
          $ 2344 "Spatula_otw" "breakAfter"
          movej(get_inverse_kin(Spatula_otw_p, qnear=Spatula_otw_q), a=1.3962634015954636, v=1.0471975511965976)
          $ 2345 "spat_S_Up_7" "breakAfter"
          movej(get_inverse_kin(spat_S_Up_7_p, qnear=spat_S_Up_7_q), a=1.3962634015954636, v=1.0471975511965976, r=0.05)
          $ 2346 "MoveL"
          $ 2347 "spat_S_Pick_4" "breakAfter"
          movel(spat_S_Pick_4_p, a=0.2, v=0.1)
          # begin: URCap Program Node
          #   Source: Robotiq_Grippers, 3.17.0.105337, Robotiq Inc.
          #   Type: Gripper
          $ 2348 "Gripper Open (1)"
          if not(gripper_connected[0]):
            popup("Gripper 1 must be connected to run this program.", "No connection", False, True, True)
          end
          if not(rq_is_gripper_activated("1")):
            popup("Gripper 1 is not activated. Go to Installation tab > Gripper to activate it and run the program again.", "Not activated", False, True, True)
          end
          rq_set_pos_spd_for(0, 255, 51, "1")
          rq_wait_pos_spe_for_request(0, 255, 51, "1")
          rq_go_to("1")
          rq_wait("1")
          # end: URCap Program Node
          $ 2349 "spat_S_Up_8" "breakAfter"
          movel(spat_S_Up_8_p, a=1.2, v=0.25, r=0.05)
          $ 2350 "Spatula_otw" "breakAfter"
          movel(Spatula_otw_p, a=1.2, v=0.25)
          $ 2351 "switch_spat_S≔ False "
          global switch_spat_S=  False
        else:
          $ 2352 "ElseIf spatula≟'spatula_flat_M'"
          if (spatula == "spatula_flat_M"):
            $ 2353 "MoveJ"
            $ 2354 "Spatula_otw" "breakAfter"
            movej(get_inverse_kin(Spatula_otw_p, qnear=Spatula_otw_q), a=1.3962634015954636, v=1.0471975511965976)
            $ 2355 "spat_flatM_up" "breakAfter"
            movej(get_inverse_kin(spat_flatM_up_p, qnear=spat_flatM_up_q), a=1.3962634015954636, v=1.0471975511965976, r=0.05)
            $ 2356 "MoveL"
            $ 2357 "spat_flatM_pick" "breakAfter"
            movel(spat_flatM_pick_p, a=0.2, v=0.1)
            # begin: URCap Program Node
            #   Source: Robotiq_Grippers, 3.17.0.105337, Robotiq Inc.
            #   Type: Gripper
            $ 2358 "Gripper Open (1)"
            if not(gripper_connected[0]):
              popup("Gripper 1 must be connected to run this program.", "No connection", False, True, True)
            end
            if not(rq_is_gripper_activated("1")):
              popup("Gripper 1 is not activated. Go to Installation tab > Gripper to activate it and run the program again.", "Not activated", False, True, True)
            end
            rq_set_pos_spd_for(0, 128, 128, "1")
            rq_wait_pos_spe_for_request(0, 128, 128, "1")
            rq_go_to("1")
            rq_wait("1")
            # end: URCap Program Node
            $ 2359 "spat_flatM_up" "breakAfter"
            movel(spat_flatM_up_p, a=1.2, v=0.25, r=0.05)
            $ 2360 "Spatula_otw" "breakAfter"
            movel(Spatula_otw_p, a=1.2, v=0.25)
            $ 2361 "switch_spat_F_M≔ False "
            global switch_spat_F_M=  False
          else:
            $ 2362 "ElseIf spatula≟'spatula_flat_S'"
            if (spatula == "spatula_flat_S"):
              $ 2363 "MoveJ"
              $ 2364 "Spatula_otw" "breakAfter"
              movej(get_inverse_kin(Spatula_otw_p, qnear=Spatula_otw_q), a=1.3962634015954636, v=1.0471975511965976)
              $ 2365 "spat_flatS_up" "breakAfter"
              movej(get_inverse_kin(spat_flatS_up_p, qnear=spat_flatS_up_q), a=1.3962634015954636, v=1.0471975511965976, r=0.05)
              $ 2366 "MoveL"
              $ 2367 "spat_flatS_pick" "breakAfter"
              movel(spat_flatS_pick_p, a=0.2, v=0.1)
              # begin: URCap Program Node
              #   Source: Robotiq_Grippers, 3.17.0.105337, Robotiq Inc.
              #   Type: Gripper
              $ 2368 "Gripper Open (1)"
              if not(gripper_connected[0]):
                popup("Gripper 1 must be connected to run this program.", "No connection", False, True, True)
              end
              if not(rq_is_gripper_activated("1")):
                popup("Gripper 1 is not activated. Go to Installation tab > Gripper to activate it and run the program again.", "Not activated", False, True, True)
              end
              rq_set_pos_spd_for(0, 128, 128, "1")
              rq_wait_pos_spe_for_request(0, 128, 128, "1")
              rq_go_to("1")
              rq_wait("1")
              # end: URCap Program Node
              $ 2369 "spat_flatS_up" "breakAfter"
              movel(spat_flatS_up_p, a=1.2, v=0.25, r=0.05)
              $ 2370 "Spatula_otw" "breakAfter"
              movel(Spatula_otw_p, a=1.2, v=0.25)
              $ 2371 "switch_spat_F_S≔ False "
              global switch_spat_F_S=  False
            end
          end
        end
      end
    end
    $ 2372 "switch_spat_M≔ True "
    global switch_spat_M=  True
    $ 2373 "switch_spat_S≔ True "
    global switch_spat_S=  True
    $ 2374 "switch_spat_F_M≔ True "
    global switch_spat_F_M=  True
    $ 2375 "switch_spat_F_S≔ True "
    global switch_spat_F_S=  True
    $ 2376 "correction_reset()"
    correction_reset()
  elif (38 == switch_1):
    $ 2572 "Case 38"
    $ 2573 "Decap Powder container"
    $ 2574 "MoveJ"
    $ 2576 "Waypoint_7" "breakAfter"
    movej(get_inverse_kin(Waypoint_7_p, qnear=Waypoint_7_q), a=1.3962634015954636, v=1.0471975511965976, r=0.05)
    $ 2577 "MoveL"
    $ 2579 "Waypoint_8" "breakAfter"
    movel(Waypoint_8_p, a=1.2, v=0.25)
    $ 2580 "MoveL"
    $ 2581 "Decapp_above_3" "breakAfter"
    movel(Decapp_above_3_p, a=1.2, v=0.25)
    $ 2582 "Set GRP_3F_Open=On"
    set_standard_digital_out(5, True)
    $ 2583 "Wait: 0.5"
    sleep(0.5)
    $ 2584 "Decapp_place_3" "breakAfter"
    movel(Decapp_place_3_p, a=0.3, v=0.05)
    $ 2585 "Set GRP_3F_Open=Off"
    set_standard_digital_out(5, False)
    $ 2586 "Wait: 0.5"
    sleep(0.5)
    # begin: URCap Program Node
    #   Source: Robotiq_Grippers, 3.17.0.105337, Robotiq Inc.
    #   Type: Gripper
    $ 2587 "Gripper Open (1)"
    if not(gripper_connected[0]):
      popup("Gripper 1 must be connected to run this program.", "No connection", False, True, True)
    end
    if not(rq_is_gripper_activated("1")):
      popup("Gripper 1 is not activated. Go to Installation tab > Gripper to activate it and run the program again.", "Not activated", False, True, True)
    end
    rq_set_pos_spd_for(0, 77, 77, "1")
    rq_wait_pos_spe_for_request(0, 77, 77, "1")
    rq_go_to("1")
    rq_wait("1")
    # end: URCap Program Node
    $ 2588 "MoveL"
    $ 2589 "Decapp_above_4" "breakAfter"
    movel(Decapp_above_4_p, a=1.2, v=0.25)
    $ 2590 "Waypoint_78" "breakAfter"
    movel(Waypoint_78_p, a=1.2, v=0.25, r=0.05)
    $ 2591 "Home (Safe)"
    movej([-1.2302089344500047, -1.2969853503591224, -1.875639182904262, -1.539621866126728, 1.5731943360401213, -2.80099559440227], a=1.3962634015954636, v=1.0471975511965976)
  elif (39 == switch_1):
    $ 2592 "Case 39"
    $ 2593 "Powder container Pick"
    $ 2594 "Direct Pick"
    $ 2595 "Set"
    set_tcp(p[0.0,0.0,0.15052000000000001,3.1415,0.0,0.0])
    $ 2596 "read_db_data()"
    read_db_data()
    # begin: URCap Program Node
    #   Source: SensoPart VISOR Robotic, 2.0.6, SensoPart Industriesensorik GmbH
    #   Type: VISOR ChangeJob
    $ 2597 "# 1 VISOR ChangeJob"
    visor_changeJob(1, "Aztec_no_dot_pick", 6000)
    # end: URCap Program Node
    # begin: URCap Program Node
    #   Source: SensoPart VISOR Robotic, 2.0.6, SensoPart Industriesensorik GmbH
    #   Type: VISOR Terminal
    $ 2598 "# 1 VISOR Terminal"
    visor_terminal(1, "TRX00", 3000)
    # end: URCap Program Node
    $ 2599 "table_pick_TCP≔visor_getPose3d(1, 0)"
    global table_pick_TCP= visor_getPose3d (1, 0)
    # begin: URCap Program Node
    #   Source: Robotiq_Grippers, 3.17.0.105337, Robotiq Inc.
    #   Type: Gripper
    $ 2600 "Gripper Open (1)"
    if not(gripper_connected[0]):
      popup("Gripper 1 must be connected to run this program.", "No connection", False, True, True)
    end
    if not(rq_is_gripper_activated("1")):
      popup("Gripper 1 is not activated. Go to Installation tab > Gripper to activate it and run the program again.", "Not activated", False, True, True)
    end
    rq_set_pos_spd_for(0, 77, 77, "1")
    rq_wait_pos_spe_for_request(0, 77, 77, "1")
    rq_go_to("1")
    rq_wait("1")
    # end: URCap Program Node
    $ 2601 "MoveJ"
    $ 2603 "Waypoint_10" "breakAfter"
    movej(get_inverse_kin(Waypoint_10_p, qnear=Waypoint_10_q), a=1.3962634015954636, v=1.0471975511965976, r=0.05)
    $ 2604 "Waypoint_9" "breakAfter"
    movej(get_inverse_kin(Waypoint_9_p, qnear=Waypoint_9_q), a=1.3962634015954636, v=1.0471975511965976, r=0.05)
    $ 2605 "MoveJ"
    $ 2607 "table_prepick≔pose_trans(table_pick_TCP,p[0,0,cent_edge/2,0,0,0])"
    global table_prepick=pose_trans(table_pick_TCP,p[0,0,cent_edge/2,0,0,0])
    $ 2608 "table_prepick" "breakAfter"
    movej(table_prepick, a=0.8726646259971648, v=0.6981317007977318)
    $ 2609 "table_safe_pick≔pose_trans(table_prepick, p[0,pick_2_base-H_c,cent_edge/2,0,0,0])"
    global table_safe_pick= pose_trans (table_prepick, p[0,pick_2_base-H_c,cent_edge/2,0,0,0])
    $ 2610 "table_safe_pick" "breakAfter"
    movej(table_safe_pick, a=0.8726646259971648, v=0.6981317007977318, r=0.05)
    $ 2611 "table_pick≔pose_trans(table_prepick, p[0,pick_2_base - d_cc,0,0,0,0])"
    global table_pick= pose_trans (table_prepick, p[0,pick_2_base - d_cc,0,0,0,0])
    $ 2612 "table_pick" "breakAfter"
    movej(table_pick, a=0.8726646259971648, v=0.6981317007977318)
    # begin: URCap Program Node
    #   Source: Robotiq_Grippers, 3.17.0.105337, Robotiq Inc.
    #   Type: Gripper
    $ 2613 "Gripper Close (1)"
    if not(gripper_connected[0]):
      popup("Gripper 1 must be connected to run this program.", "No connection", False, True, True)
    end
    if not(rq_is_gripper_activated("1")):
      popup("Gripper 1 is not activated. Go to Installation tab > Gripper to activate it and run the program again.", "Not activated", False, True, True)
    end
    rq_set_pos_spd_for(255, 77, 51, "1")
    rq_wait_pos_spe_for_request(255, 77, 51, "1")
    rq_go_to("1")
    rq_wait("1")
    # end: URCap Program Node
    $ 2614 "table_prepick" "breakAfter"
    movej(table_prepick, a=0.8726646259971648, v=0.6981317007977318)
    $ 2615 "Picking≔ True "
    global Picking=  True
    $ 2617 "powder_position≔'Position2'"
    global powder_position="Position2"
    $ 2618 "MoveJ"
    $ 2619 "Powder_wayp1" "breakAfter"
    movej(get_inverse_kin(Powder_wayp1_p, qnear=Powder_wayp1_q), a=1.3962634015954636, v=1.0471975511965976, r=0.05)
    $ 2620 "MoveL"
    $ 2621 "Waypoint_2" "breakAfter"
    movel(Waypoint_2_p, a=1.2, v=0.25)
    $ 2622 "Set"
    set_tcp(p[0.0,0.0,0.161,3.1415,0.0,0.0])
    $ 2623 "If powder_position ≟ 'Position1'"
    if (powder_position  ==  "Position1"):
      $ 2624 "MoveJ"
      $ 2625 "Postions_otw" "breakAfter"
      movej(get_inverse_kin(Postions_otw_p, qnear=Postions_otw_q), a=1.3962634015954636, v=1.0471975511965976, r=0.01)
      $ 2626 "MoveL"
      $ 2627 "Cont_A_TCP" "breakAfter"
      movel(Cont_A_TCP, a=0.5, v=0.2)
      $ 2628 "cont_A_prepick≔pose_trans(Cont_A_TCP, p[0,0,cent_edge/2,0,0,0])"
      global cont_A_prepick= pose_trans (Cont_A_TCP, p[0,0,cent_edge/2,0,0,0])
      $ 2629 "cont_A_prepick" "breakAfter"
      movel(cont_A_prepick, a=0.3, v=0.05)
      $ 2630 "cont_A_pick≔pose_trans(cont_A_prepick, p[0,pick_2_base-d_cc,0,0,0,0])"
      global cont_A_pick= pose_trans (cont_A_prepick, p[0,pick_2_base-d_cc,0,0,0,0])
      $ 2631 "cont_A_pick" "breakAfter"
      movel(cont_A_pick, a=0.2, v=0.1)
      # begin: URCap Program Node
      #   Source: Robotiq_Grippers, 3.17.0.105337, Robotiq Inc.
      #   Type: Gripper
      $ 2632 "Gripper Open (1)"
      if not(gripper_connected[0]):
        popup("Gripper 1 must be connected to run this program.", "No connection", False, True, True)
      end
      if not(rq_is_gripper_activated("1")):
        popup("Gripper 1 is not activated. Go to Installation tab > Gripper to activate it and run the program again.", "Not activated", False, True, True)
      end
      rq_set_pos_spd_for(0, 77, 26, "1")
      rq_wait_pos_spe_for_request(0, 77, 26, "1")
      rq_go_to("1")
      rq_wait("1")
      # end: URCap Program Node
      $ 2633 "cont_A_otw" "breakAfter"
      movel(cont_A_otw_p, a=0.5, v=0.2)
      $ 2634 "cont_A_prepick" "breakAfter"
      movel(cont_A_prepick, a=0.5, v=0.2)
      $ 2635 "Postions_otw" "breakAfter"
      movel(Postions_otw_p, a=0.5, v=0.2, r=0.01)
      $ 2637 "Home (Safe)"
      movej([-1.2302089344500047, -1.2969853503591224, -1.875639182904262, -1.539621866126728, 1.5731943360401213, -2.80099559440227], a=1.3962634015954636, v=1.0471975511965976)
    else:
      $ 2639 "ElseIf powder_position≟'Position2'"
      if (powder_position == "Position2"):
        $ 2640 "MoveJ"
        $ 2641 "Postions_otw" "breakAfter"
        movej(get_inverse_kin(Postions_otw_p, qnear=Postions_otw_q), a=1.3962634015954636, v=1.0471975511965976, r=0.01)
        $ 2642 "MoveL"
        $ 2645 "cont_B_prepick≔pose_trans(Cont_B_TCP, p[0,0,cent_edge/2,0,0,0])"
        global cont_B_prepick= pose_trans (Cont_B_TCP, p[0,0,cent_edge/2,0,0,0])
        $ 2646 "cont_B_prepick" "breakAfter"
        movel(cont_B_prepick, a=1.2, v=0.25)
        $ 2647 "cont_B_pick≔pose_trans(cont_B_prepick, p[0,pick_2_base-d_cc,0,0,0,0])"
        global cont_B_pick= pose_trans (cont_B_prepick, p[0,pick_2_base-d_cc,0,0,0,0])
        $ 2648 "cont_B_pick" "breakAfter"
        global move_thread_flag_2648=0
        thread move_thread_2648():
          enter_critical
          move_thread_flag_2648 = 1
          movel(cont_B_pick, a=0.2, v=0.1)
          move_thread_flag_2648 = 2
          exit_critical
        end
        move_thread_flag_2648 = 0
        move_thread_han_2648 = run move_thread_2648()
        while (True):
          local targetTcpDirection=get_target_tcp_speed()
          local stepsToRetract=tool_contact(direction=targetTcpDirection, force_threshold=8.000000)
          if (stepsToRetract > 0):
            kill move_thread_han_2648
            stopl(3.0)
            local backTrackMovement=get_actual_joint_positions_history(stepsToRetract)
            local contactPose=get_forward_kin(backTrackMovement)
            local posDir=[targetTcpDirection[0],targetTcpDirection[1],targetTcpDirection[2]]
            local retractTo=contactPose
            if (norm(posDir) > 1e-6):
              local normalizedPosDir=normalize(posDir)
              local additionalRetraction=p[normalizedPosDir[0] * 0.0, normalizedPosDir[1] * 0.0, normalizedPosDir[2] * 0.0, 0, 0, 0]
              retractTo = pose_sub(contactPose, additionalRetraction)
            end
            movel(retractTo, a=3.0, v=0.1)
            $ 2649 "Until (tool_contact_detection)"
            $ 2650 "saved_place_pos≔get_actual_tcp_pose()"
            global saved_place_pos= get_actual_tcp_pose ()
            break
          end
          sleep(1.0E-10)
          if (move_thread_flag_2648 > 1):
            join move_thread_han_2648
            break
          end
          sync()
        end
        # begin: URCap Program Node
        #   Source: Robotiq_Grippers, 3.17.0.105337, Robotiq Inc.
        #   Type: Gripper
        $ 2651 "Gripper Open (1)"
        if not(gripper_connected[0]):
          popup("Gripper 1 must be connected to run this program.", "No connection", False, True, True)
        end
        if not(rq_is_gripper_activated("1")):
          popup("Gripper 1 is not activated. Go to Installation tab > Gripper to activate it and run the program again.", "Not activated", False, True, True)
        end
        rq_set_pos_spd_for(0, 77, 26, "1")
        rq_wait_pos_spe_for_request(0, 77, 26, "1")
        rq_go_to("1")
        rq_wait("1")
        # end: URCap Program Node
        $ 2652 "cont_B_otw" "breakAfter"
        movel(cont_B_otw_p, a=1.2, v=0.25)
        $ 2654 "cont_B_safe" "breakAfter"
        movel(cont_B_safe_p, a=1.2, v=0.25)
        $ 2655 "Postions_otw" "breakAfter"
        movel(Postions_otw_p, a=1.2, v=0.25)
        $ 2656 "Home (Safe)"
        movej([-1.2302089344500047, -1.2969853503591224, -1.875639182904262, -1.539621866126728, 1.5731943360401213, -2.80099559440227], a=1.3962634015954636, v=1.0471975511965976)
      else:
        $ 2658 "ElseIf powder_position≟'Position3'"
        if (powder_position == "Position3"):
          $ 2659 "MoveJ"
          $ 2660 "Postions_otw" "breakAfter"
          movej(get_inverse_kin(Postions_otw_p, qnear=Postions_otw_q), a=1.3962634015954636, v=1.0471975511965976, r=0.01)
          $ 2667 "MoveL"
          $ 2668 "Cont_C_TCP" "breakAfter"
          movel(Cont_C_TCP, a=1.2, v=0.25, r=0.01)
          $ 2669 "cont_C_prepick≔pose_trans(Cont_C_TCP, p[0,0,cent_edge/2,0,0,0])"
          global cont_C_prepick= pose_trans (Cont_C_TCP, p[0,0,cent_edge/2,0,0,0])
          $ 2670 "cont_C_prepick" "breakAfter"
          movel(cont_C_prepick, a=0.3, v=0.05)
          $ 2671 "cont_C_pick≔pose_trans(cont_C_prepick, p[0,pick_2_base-d_cc,0,0,0,0])"
          global cont_C_pick= pose_trans (cont_C_prepick, p[0,pick_2_base-d_cc,0,0,0,0])
          $ 2672 "cont_C_pick" "breakAfter"
          movel(cont_C_pick, a=0.2, v=0.1)
          # begin: URCap Program Node
          #   Source: Robotiq_Grippers, 3.17.0.105337, Robotiq Inc.
          #   Type: Gripper
          $ 2673 "Gripper Open (1)"
          if not(gripper_connected[0]):
            popup("Gripper 1 must be connected to run this program.", "No connection", False, True, True)
          end
          if not(rq_is_gripper_activated("1")):
            popup("Gripper 1 is not activated. Go to Installation tab > Gripper to activate it and run the program again.", "Not activated", False, True, True)
          end
          rq_set_pos_spd_for(0, 77, 26, "1")
          rq_wait_pos_spe_for_request(0, 77, 26, "1")
          rq_go_to("1")
          rq_wait("1")
          # end: URCap Program Node
          $ 2674 "cont_C_otw" "breakAfter"
          movel(cont_C_otw_p, a=1.2, v=0.25)
          $ 2675 "cont_C_prepick" "breakAfter"
          movel(cont_C_prepick, a=1.2, v=0.25, r=0.01)
          $ 2676 "Postions_otw" "breakAfter"
          movel(Postions_otw_p, a=1.2, v=0.25)
          $ 2677 "Home (Safe)"
          movej([-1.2302089344500047, -1.2969853503591224, -1.875639182904262, -1.539621866126728, 1.5731943360401213, -2.80099559440227], a=1.3962634015954636, v=1.0471975511965976)
        end
      end
    end
    $ 2679 "Home (Safe)"
    movej([-1.2302089344500047, -1.2969853503591224, -1.875639182904262, -1.539621866126728, 1.5731943360401213, -2.80099559440227], a=1.3962634015954636, v=1.0471975511965976)
  elif (41 == switch_1):
    $ 2788 "Case 41"
    $ 2789 "Task≔'Decapping_Dosing'"
    global Task="Decapping_Dosing"
    $ 2790 "tilt_to_home()"
    tilt_to_home()
    $ 2791 "Weigh, Place & decap container"
    $ 2792 "Set"
    set_tcp(p[0.0,0.0,0.15052000000000001,3.1415,0.0,0.0])
    # begin: URCap Program Node
    #   Source: SensoPart VISOR Robotic, 2.0.6, SensoPart Industriesensorik GmbH
    #   Type: VISOR Robotic App
    $ 2793 "VISOR Easy Pick"
    def visorFuncEasyPick_47a8ba():
      # begin: URCap Program Node
      #   Source: SensoPart VISOR Robotic, 2.0.6, SensoPart Industriesensorik GmbH
      #   Type: Easy Pick Setup
      $ 2794 "# 1 Setup" "noBreak"
      local easyPickVisorId = 1
      local easyPickArmMounted = True
      local easyPickSetJob = True
      local easyPickJobName = "PoTS"
      local easyPickAtImgAcq = False
      local easyPickImgAcqPose = FRM_PoTS
      # end: URCap Program Node
      # begin: URCap Program Node
      #   Source: SensoPart VISOR Robotic, 2.0.6, SensoPart Industriesensorik GmbH
      #   Type: Process
      $ 2795 "Process" "noBreak"
      local easyPickObjTaken = False
      local easyPickTrigger = False
      local easyPickPoseIdx = 0
      local easyPickPose = p[0,0,0,0,0,0]
      def easyPickFuncTrigger(visorId, setJob, jobName, arm):
      if (setJob):
        visor_changeJob(visorId, jobName, 6000)
      end
      if (arm):
        visor_trigger(visorId, 6000, "arm")
      else:
        visor_trigger(visorId, 6000)
      end
      global easyPickParts_7=visor_partsFound(visorId)
      visor_easyPickUpdate(visorId, "parts", visor_partsFound(visorId))
      return visor_getPose3d(visorId, 0)
    end
    while (not easyPickObjTaken):
      easyPickTrigger = (easyPickCount_7 >= visor_partsFound(easyPickVisorId)) or (easyPickCount_7 > 9) or (not visor_easyPickCheckIdent("d8ba5f", easyPickVisorId))
      if (easyPickTrigger):
        easyPickCount_7 = 0
      end
      easyPickPoseIdx = easyPickCount_7
      easyPickPose = visor_getPose3d(easyPickVisorId, easyPickPoseIdx)
      visor_easyPickUpdate(easyPickVisorId, "counter", easyPickPoseIdx)
      # begin: URCap Program Node
      #   Source: SensoPart VISOR Robotic, 2.0.6, SensoPart Industriesensorik GmbH
      #   Type: Image Acquisition Pose
      $ 2796 "Image Acquisition Pose" "noBreak"
      if (easyPickTrigger):
        if (not easyPickAtImgAcq):
          movej(pose_trans(easyPickImgAcqPose,p[0.0000,0.0000,-0.0000,0.0000,0.0000,0.0000]),a=1.3963,v=1.0472,t=0.000000,r=0.000000)
          easyPickAtImgAcq = True
        end
        easyPickPose = easyPickFuncTrigger(easyPickVisorId, easyPickSetJob, easyPickJobName, easyPickArmMounted)
      end
      # end: URCap Program Node
      # begin: URCap Program Node
      #   Source: SensoPart VISOR Robotic, 2.0.6, SensoPart Industriesensorik GmbH
      #   Type: Object Detected
      $ 2797 "Object Detected" "noBreak"
      if (visor_partsFound(easyPickVisorId) > 0):
        $ 2798 "Open Gripper" "noBreak"
        # begin: URCap Program Node
        #   Source: Robotiq_Grippers, 3.17.0.105337, Robotiq Inc.
        #   Type: Gripper
        $ 2799 "Gripper Open (1)" "noBreak"
        if not(gripper_connected[0]):
          popup("Gripper 1 must be connected to run this program.", "No connection", False, True, True)
        end
        if not(rq_is_gripper_activated("1")):
          popup("Gripper 1 is not activated. Go to Installation tab > Gripper to activate it and run the program again.", "Not activated", False, True, True)
        end
        rq_set_pos_spd_for(0, 77, 77, "1")
        rq_wait_pos_spe_for_request(0, 77, 77, "1")
        rq_go_to("1")
        rq_wait("1")
        # end: URCap Program Node
        $ 2800 "Set" "noBreak"
        set_tcp(p[0.0,0.0,0.161,3.1415,0.0,0.0])
        $ 2801 "Wait: 0.2" "noBreak"
        sleep(0.2)
        $ 2802 "Place on second weigh scale" "noBreak"
        $ 2803 "MoveJ" "noBreak"
        $ 2804 "Waypoint_1" "noBreak"
        movej(get_inverse_kin(Waypoint_1_p, qnear=Waypoint_1_q), a=1.3962634015954636, v=1.0471975511965976, r=0.1)
        $ 2805 "Waypoint_5" "noBreak"
        movej(get_inverse_kin(Waypoint_5_p, qnear=Waypoint_5_q), a=1.3962634015954636, v=1.0471975511965976)
        $ 2807 "If Picking≟ True " "noBreak"
        if (Picking ==   True  ):
          $ 2808 "Pick from saved pose" "noBreak"
          $ 2809 "MoveL" "noBreak"
          $ 2810 "cont_B_safe" "noBreak"
          movel(cont_B_safe_p, a=0.2, v=0.1)
          $ 2811 "saved_place_pos" "noBreak"
          movel(saved_place_pos, a=1.2, v=0.25)
          # begin: URCap Program Node
          #   Source: Robotiq_Grippers, 3.17.0.105337, Robotiq Inc.
          #   Type: Gripper
          $ 2812 "Gripper Close (1)" "noBreak"
          if not(gripper_connected[0]):
            popup("Gripper 1 must be connected to run this program.", "No connection", False, True, True)
          end
          if not(rq_is_gripper_activated("1")):
            popup("Gripper 1 is not activated. Go to Installation tab > Gripper to activate it and run the program again.", "Not activated", False, True, True)
          end
          rq_set_pos_spd_for(255, 77, 26, "1")
          rq_wait_pos_spe_for_request(255, 77, 26, "1")
          rq_go_to("1")
          rq_wait("1")
          # end: URCap Program Node
          $ 2813 "cont_B_safe" "noBreak"
          movel(cont_B_safe_p, a=1.2, v=0.25)
          $ 2814 "Postions_otw" "noBreak"
          movel(Postions_otw_p, a=1.2, v=0.25)
        else:
          $ 2817 "Else" "noBreak"
          $ 2818 "read_db_data()" "noBreak"
          read_db_data()
          $ 2819 "Pick from B" "noBreak"
          $ 2820 "MoveL" "noBreak"
          $ 2822 "cont_B_safe" "noBreak"
          movel(cont_B_safe_p, a=1.2, v=0.25)
          $ 2823 "cont_B_prepick≔pose_trans(Cont_B_TCP, p[0,0,cent_edge/2,0,0,0])" "noBreak"
          global cont_B_prepick= pose_trans (Cont_B_TCP, p[0,0,cent_edge/2,0,0,0])
          $ 2824 "cont_B_otw" "noBreak"
          movel(cont_B_otw_p, a=1.2, v=0.25)
          $ 2826 "cont_B_pick≔pose_trans(cont_B_prepick, p[0,pick_2_base-d_cc,0,0,0,0])" "noBreak"
          global cont_B_pick= pose_trans (cont_B_prepick, p[0,pick_2_base-d_cc,0,0,0,0])
          $ 2827 "cont_B_pick" "noBreak"
          movel(cont_B_pick, a=0.2, v=0.1)
          # begin: URCap Program Node
          #   Source: Robotiq_Grippers, 3.17.0.105337, Robotiq Inc.
          #   Type: Gripper
          $ 2828 "Gripper Close (1)" "noBreak"
          if not(gripper_connected[0]):
            popup("Gripper 1 must be connected to run this program.", "No connection", False, True, True)
          end
          if not(rq_is_gripper_activated("1")):
            popup("Gripper 1 is not activated. Go to Installation tab > Gripper to activate it and run the program again.", "Not activated", False, True, True)
          end
          rq_set_pos_spd_for(255, 77, 51, "1")
          rq_wait_pos_spe_for_request(255, 77, 51, "1")
          rq_go_to("1")
          rq_wait("1")
          # end: URCap Program Node
          $ 2829 "cont_B_prepick" "noBreak"
          movel(cont_B_prepick, a=1.2, v=0.25, r=0.01)
          $ 2830 "Postions_otw" "noBreak"
          movel(Postions_otw_p, a=1.2, v=0.25)
        end
        $ 2847 "Set" "noBreak"
        set_tcp(p[0.0,0.0,0.15052000000000001,3.1415,0.0,0.0])
        # begin: URCap Program Node
        #   Source: SensoPart VISOR Robotic, 2.0.6, SensoPart Industriesensorik GmbH
        #   Type: Approach Pose
        $ 2848 "Approach Pose" "noBreak"
        movej(pose_trans(easyPickPose,p[0.0000,0.0000,-0.0000,0.0000,0.0000,0.0000]),a=0.5236,v=0.4363,t=0.000000,r=0.000000)
        # end: URCap Program Node
        # begin: URCap Program Node
        #   Source: SensoPart VISOR Robotic, 2.0.6, SensoPart Industriesensorik GmbH
        #   Type: Target Pose
        $ 2849 "Target Pose" "noBreak"
        movel(pose_trans(easyPickPose,p[0.0000,0.0000,-0.0000,0.0000,0.0000,0.0000]),a=0.1000,v=0.0500,t=0.000000,r=0.000000)
        # end: URCap Program Node
        $ 2850 "Close Gripper" "noBreak"
        $ 2851 "container_place≔get_actual_tcp_pose()" "noBreak"
        global container_place= get_actual_tcp_pose ()
        $ 2852 "PoTS_place_abov≔pose_trans(container_place, p[0,0,cent_edge/2,0,0,0])" "noBreak"
        global PoTS_place_abov=pose_trans(container_place, p[0,0,cent_edge/2,0,0,0])
        $ 2853 "MoveL" "noBreak"
        $ 2854 "PoTS_place_abov" "noBreak"
        movel(PoTS_place_abov, a=0.5, v=0.05)
        $ 2856 "target_pose≔pose_trans(PoTS_place_abov, p[0,pick_2_base-d_cc,0,0,0,0])" "noBreak"
        global target_pose=pose_trans(PoTS_place_abov, p[0,pick_2_base-d_cc,0,0,0,0])
        $ 2857 "MoveL" "noBreak"
        $ 2858 "target_pose" "noBreak"
        movel(target_pose, a=0.3, v=0.05)
        # begin: URCap Program Node
        #   Source: Robotiq_Grippers, 3.17.0.105337, Robotiq Inc.
        #   Type: Gripper
        $ 2859 "Gripper Open (1)" "noBreak"
        if not(gripper_connected[0]):
          popup("Gripper 1 must be connected to run this program.", "No connection", False, True, True)
        end
        if not(rq_is_gripper_activated("1")):
          popup("Gripper 1 is not activated. Go to Installation tab > Gripper to activate it and run the program again.", "Not activated", False, True, True)
        end
        rq_set_pos_spd_for(0, 77, 77, "1")
        rq_wait_pos_spe_for_request(0, 77, 77, "1")
        rq_go_to("1")
        rq_wait("1")
        # end: URCap Program Node
        # begin: URCap Program Node
        #   Source: SensoPart VISOR Robotic, 2.0.6, SensoPart Industriesensorik GmbH
        #   Type: Exit Pose
        $ 2860 "Exit Pose" "noBreak"
        movel(pose_trans(easyPickPose,p[0.0000,0.0000,0.1000,0.0000,0.0000,0.0000]),a=0.5000,v=0.2500,t=0.000000,r=0.000000)
        # end: URCap Program Node
        easyPickObjTaken = True
      end
      # end: URCap Program Node
      # begin: URCap Program Node
      #   Source: SensoPart VISOR Robotic, 2.0.6, SensoPart Industriesensorik GmbH
      #   Type: No Object Detected
      $ 2861 "No Object Detected" "noBreak"
      if (visor_partsFound(easyPickVisorId) < 1):
        $ 2862 "Popup: No POTS detected" "noBreak"
        popup("No POTS detected", "Message", False, False, blocking=True)
        else:
      end
      # end: URCap Program Node
    end
    easyPickCount_7 = easyPickCount_7 + 1
    visor_easyPickUpdate(easyPickVisorId, "counter", easyPickCount_7)
    visor_easyPickSetIdent("d8ba5f", easyPickVisorId)
    # end: URCap Program Node
  end
  visorFuncEasyPick_47a8ba()
  # end: URCap Program Node
  $ 2897 "MoveJ"
  $ 2898 "place_2_home" "breakAfter"
  movej(get_inverse_kin(place_2_home_p, qnear=place_2_home_q), a=1.3962634015954636, v=1.0471975511965976)
  $ 2899 "Picking≔ False "
  global Picking=  False
  elif (42 == switch_1):
    $ 2900 "Case 42"
  elif (43 == switch_1):
    $ 3662 "Case 43"
  elif (44 == switch_1):
    $ 3915 "Case 44"
  elif (45 == switch_1):
    $ 3979 "Case 45"
  elif (46 == switch_1):
    $ 4016 "Case 46"
  elif (47 == switch_1):
    $ 4306 "Case 47"
  elif (48 == switch_1):
    $ 4361 "Case 48"
  elif (49 == switch_1):
    $ 4379 "Case 49"
  elif (50 == switch_1):
    $ 4397 "Case 50"
    $ 4398 "Emptying powder container"
    $ 4399 "tilt_to_home()"
    tilt_to_home()
    $ 4400 "scoop_status≔'emptying'"
    global scoop_status="emptying"
    $ 4401 "Dosing untill empty"
    $ 4402 "tilt_angle_sent≔0.0"
    global tilt_angle_sent=0.0
    $ 4403 "send_target_info()"
    send_target_info()
    $ 4404 "zero_scale()"
    zero_scale()
    $ 4405 "prev_spat≔''"
    global prev_spat=""
    $ 4406 "spatula≔''"
    global spatula=""
    $ 4407 "send_powder_info()"
    send_powder_info()
    $ 4408 "Set AO[0]=0.0"
    set_standard_analog_out(0, 0.0)
    $ 4409 "Wait: 0.2"
    sleep(0.2)
    $ 4410 "reach pots decapping pose"
    # begin: URCap Program Node
    #   Source: SensoPart VISOR Robotic, 2.0.6, SensoPart Industriesensorik GmbH
    #   Type: VISOR Robotic App
    $ 4416 "VISOR Easy Pick"
    def visorFuncEasyPick_8737ac():
      # begin: URCap Program Node
      #   Source: SensoPart VISOR Robotic, 2.0.6, SensoPart Industriesensorik GmbH
      #   Type: Easy Pick Setup
      $ 4417 "# 1 Setup" "noBreak"
      local easyPickVisorId = 1
      local easyPickArmMounted = True
      local easyPickSetJob = True
      local easyPickJobName = "Weight_scale"
      local easyPickAtImgAcq = False
      local easyPickImgAcqPose = Trigger
      # end: URCap Program Node
      # begin: URCap Program Node
      #   Source: SensoPart VISOR Robotic, 2.0.6, SensoPart Industriesensorik GmbH
      #   Type: Process
      $ 4418 "Process" "noBreak"
      local easyPickObjTaken = False
      local easyPickTrigger = False
      local easyPickPoseIdx = 0
      local easyPickPose = p[0,0,0,0,0,0]
      def easyPickFuncTrigger(visorId, setJob, jobName, arm):
      if (setJob):
        visor_changeJob(visorId, jobName, 6000)
      end
      if (arm):
        visor_trigger(visorId, 6000, "arm")
      else:
        visor_trigger(visorId, 6000)
      end
      global easyPickParts_4=visor_partsFound(visorId)
      visor_easyPickUpdate(visorId, "parts", visor_partsFound(visorId))
      return visor_getPose3d(visorId, 0)
    end
    while (not easyPickObjTaken):
      easyPickTrigger = (easyPickCount_4 >= visor_partsFound(easyPickVisorId)) or (easyPickCount_4 > 9) or (not visor_easyPickCheckIdent("bfde9f", easyPickVisorId))
      if (easyPickTrigger):
        easyPickCount_4 = 0
      end
      easyPickPoseIdx = easyPickCount_4
      easyPickPose = visor_getPose3d(easyPickVisorId, easyPickPoseIdx)
      visor_easyPickUpdate(easyPickVisorId, "counter", easyPickPoseIdx)
      # begin: URCap Program Node
      #   Source: SensoPart VISOR Robotic, 2.0.6, SensoPart Industriesensorik GmbH
      #   Type: Image Acquisition Pose
      $ 4419 "Image Acquisition Pose" "noBreak"
      if (easyPickTrigger):
        if (not easyPickAtImgAcq):
          movej(pose_trans(easyPickImgAcqPose,p[0.0000,0.0000,-0.0000,0.0000,0.0000,0.0000]),a=1.3963,v=1.0472,t=0.000000,r=0.000000)
          easyPickAtImgAcq = True
        end
        easyPickPose = easyPickFuncTrigger(easyPickVisorId, easyPickSetJob, easyPickJobName, easyPickArmMounted)
      end
      # end: URCap Program Node
      # begin: URCap Program Node
      #   Source: SensoPart VISOR Robotic, 2.0.6, SensoPart Industriesensorik GmbH
      #   Type: Object Detected
      $ 4420 "Object Detected" "noBreak"
      if (visor_partsFound(easyPickVisorId) > 0):
        $ 4421 "Open Gripper" "noBreak"
        $ 4422 "weight_value≔get_weight()" "noBreak"
        global weight_value=get_weight()
        $ 4423 "Wait: 1.0" "noBreak"
        sleep(1.0)
        $ 4424 "diff≔target_weight-weight_value" "noBreak"
        global diff=target_weight-weight_value
        $ 4425 "compute_level_percent(W_now, weight_value)" "noBreak"
        compute_level_percent(W_now, weight_value)
        $ 4426 "send_level_info()" "noBreak"
        send_level_info()
        $ 4427 "spatula≔select_spatula(Flowability, level, diff, bulk_density, mouth_d)" "noBreak"
        global spatula=select_spatula(Flowability, level, diff, bulk_density, mouth_d)
        $ 4428 "Wait: 0.2" "noBreak"
        sleep(0.2)
        $ 4429 "send_spatula_info()" "noBreak"
        send_spatula_info()
        $ 4430 "Pick spatula" "noBreak"
        $ 4431 "If spatula ≟ 'spatula_L'" "noBreak"
        if (spatula  ==  "spatula_L"):
          $ 4432 "MoveJ" "noBreak"
          $ 4433 "Spatula_otw" "noBreak"
          movej(get_inverse_kin(Spatula_otw_p, qnear=Spatula_otw_q), a=1.3962634015954636, v=1.0471975511965976)
          $ 4434 "pick_spat_L_abv" "noBreak"
          movej(get_inverse_kin(pick_spat_L_abv_p, qnear=pick_spat_L_abv_q), a=1.3962634015954636, v=1.0471975511965976)
          $ 4435 "MoveL" "noBreak"
          $ 4436 "spat_L_pick" "noBreak"
          movel(spat_L_pick_p, a=1.2, v=0.25)
          # begin: URCap Program Node
          #   Source: Robotiq_Grippers, 3.17.0.105337, Robotiq Inc.
          #   Type: Gripper
          $ 4437 "Gripper Close (1)" "noBreak"
          if not(gripper_connected[0]):
            popup("Gripper 1 must be connected to run this program.", "No connection", False, True, True)
          end
          if not(rq_is_gripper_activated("1")):
            popup("Gripper 1 is not activated. Go to Installation tab > Gripper to activate it and run the program again.", "Not activated", False, True, True)
          end
          rq_set_pos_spd_for(255, 0, 77, "1")
          rq_wait_pos_spe_for_request(255, 0, 77, "1")
          rq_go_to("1")
          rq_wait("1")
          # end: URCap Program Node
          $ 4438 "spat_L_lift" "noBreak"
          movel(spat_L_lift_p, a=1.2, v=0.25, r=0.01)
          $ 4439 "spat_L_side" "noBreak"
          movel(spat_L_side_p, a=1.2, v=0.25, r=0.01)
          $ 4440 "spat_L_up" "noBreak"
          movel(spat_L_up_p, a=1.2, v=0.25, r=0.05)
          $ 4441 "MoveJ" "noBreak"
          $ 4442 "Spatula_otw" "noBreak"
          movej(get_inverse_kin(Spatula_otw_p, qnear=Spatula_otw_q), a=1.3962634015954636, v=1.0471975511965976)
        else:
          $ 4443 "ElseIf spatula ≟'spatula_M'" "noBreak"
          if (spatula  == "spatula_M"):
            $ 4444 "MoveJ" "noBreak"
            $ 4445 "Spatula_otw" "noBreak"
            movej(get_inverse_kin(Spatula_otw_p, qnear=Spatula_otw_q), a=1.3962634015954636, v=1.0471975511965976)
            $ 4446 "spat_M_up" "noBreak"
            movej(get_inverse_kin(spat_M_up_p, qnear=spat_M_up_q), a=1.3962634015954636, v=1.0471975511965976, r=0.05)
            $ 4447 "MoveL" "noBreak"
            $ 4448 "spat_M_pick" "noBreak"
            movel(spat_M_pick_p, a=1.2, v=0.25)
            # begin: URCap Program Node
            #   Source: Robotiq_Grippers, 3.17.0.105337, Robotiq Inc.
            #   Type: Gripper
            $ 4449 "Gripper Close (1)" "noBreak"
            if not(gripper_connected[0]):
              popup("Gripper 1 must be connected to run this program.", "No connection", False, True, True)
            end
            if not(rq_is_gripper_activated("1")):
              popup("Gripper 1 is not activated. Go to Installation tab > Gripper to activate it and run the program again.", "Not activated", False, True, True)
            end
            rq_set_pos_spd_for(255, 0, 77, "1")
            rq_wait_pos_spe_for_request(255, 0, 77, "1")
            rq_go_to("1")
            rq_wait("1")
            # end: URCap Program Node
            $ 4450 "spat_M_up" "noBreak"
            movel(spat_M_up_p, a=1.2, v=0.25, r=0.05)
            $ 4451 "Spatula_otw" "noBreak"
            movel(Spatula_otw_p, a=1.2, v=0.25)
            $ 4452 "switch_spat_M≔ False " "noBreak"
            global switch_spat_M=  False
          else:
            $ 4453 "ElseIf spatula≟'spatula_S'" "noBreak"
            if (spatula == "spatula_S"):
              $ 4454 "MoveJ" "noBreak"
              $ 4455 "Spatula_otw" "noBreak"
              movej(get_inverse_kin(Spatula_otw_p, qnear=Spatula_otw_q), a=1.3962634015954636, v=1.0471975511965976)
              $ 4456 "spat_S_Up_7" "noBreak"
              movej(get_inverse_kin(spat_S_Up_7_p, qnear=spat_S_Up_7_q), a=1.3962634015954636, v=1.0471975511965976, r=0.05)
              $ 4457 "MoveL" "noBreak"
              $ 4458 "spat_S_Pick_4" "noBreak"
              movel(spat_S_Pick_4_p, a=1.2, v=0.25)
              # begin: URCap Program Node
              #   Source: Robotiq_Grippers, 3.17.0.105337, Robotiq Inc.
              #   Type: Gripper
              $ 4459 "Gripper Close (1)" "noBreak"
              if not(gripper_connected[0]):
                popup("Gripper 1 must be connected to run this program.", "No connection", False, True, True)
              end
              if not(rq_is_gripper_activated("1")):
                popup("Gripper 1 is not activated. Go to Installation tab > Gripper to activate it and run the program again.", "Not activated", False, True, True)
              end
              rq_set_pos_spd_for(255, 0, 77, "1")
              rq_wait_pos_spe_for_request(255, 0, 77, "1")
              rq_go_to("1")
              rq_wait("1")
              # end: URCap Program Node
              $ 4460 "spat_S_Up_8" "noBreak"
              movel(spat_S_Up_8_p, a=1.2, v=0.25, r=0.05)
              $ 4461 "Spatula_otw" "noBreak"
              movel(Spatula_otw_p, a=1.2, v=0.25)
              $ 4462 "switch_spat_S≔ False " "noBreak"
              global switch_spat_S=  False
            else:
              $ 4463 "ElseIf spatula≟'spatula_flat_M'" "noBreak"
              if (spatula == "spatula_flat_M"):
                $ 4464 "MoveJ" "noBreak"
                $ 4465 "Spatula_otw" "noBreak"
                movej(get_inverse_kin(Spatula_otw_p, qnear=Spatula_otw_q), a=1.3962634015954636, v=1.0471975511965976)
                $ 4466 "spat_flatM_up" "noBreak"
                movej(get_inverse_kin(spat_flatM_up_p, qnear=spat_flatM_up_q), a=1.3962634015954636, v=1.0471975511965976, r=0.05)
                $ 4467 "MoveL" "noBreak"
                $ 4468 "spat_flatM_pick" "noBreak"
                movel(spat_flatM_pick_p, a=1.2, v=0.25)
                # begin: URCap Program Node
                #   Source: Robotiq_Grippers, 3.17.0.105337, Robotiq Inc.
                #   Type: Gripper
                $ 4469 "Gripper Close (1)" "noBreak"
                if not(gripper_connected[0]):
                  popup("Gripper 1 must be connected to run this program.", "No connection", False, True, True)
                end
                if not(rq_is_gripper_activated("1")):
                  popup("Gripper 1 is not activated. Go to Installation tab > Gripper to activate it and run the program again.", "Not activated", False, True, True)
                end
                rq_set_pos_spd_for(255, 0, 77, "1")
                rq_wait_pos_spe_for_request(255, 0, 77, "1")
                rq_go_to("1")
                rq_wait("1")
                # end: URCap Program Node
                $ 4470 "spat_flatM_up" "noBreak"
                movel(spat_flatM_up_p, a=1.2, v=0.25, r=0.05)
                $ 4471 "Spatula_otw" "noBreak"
                movel(Spatula_otw_p, a=1.2, v=0.25)
                $ 4472 "switch_spat_F_M≔ False " "noBreak"
                global switch_spat_F_M=  False
              else:
                $ 4473 "ElseIf spatula≟'spatula_flat_S'" "noBreak"
                if (spatula == "spatula_flat_S"):
                  $ 4474 "MoveJ" "noBreak"
                  $ 4475 "Spatula_otw" "noBreak"
                  movej(get_inverse_kin(Spatula_otw_p, qnear=Spatula_otw_q), a=1.3962634015954636, v=1.0471975511965976)
                  $ 4476 "spat_flatS_up" "noBreak"
                  movej(get_inverse_kin(spat_flatS_up_p, qnear=spat_flatS_up_q), a=1.3962634015954636, v=1.0471975511965976, r=0.05)
                  $ 4477 "MoveL" "noBreak"
                  $ 4478 "spat_flatS_pick" "noBreak"
                  movel(spat_flatS_pick_p, a=1.2, v=0.25)
                  # begin: URCap Program Node
                  #   Source: Robotiq_Grippers, 3.17.0.105337, Robotiq Inc.
                  #   Type: Gripper
                  $ 4479 "Gripper Close (1)" "noBreak"
                  if not(gripper_connected[0]):
                    popup("Gripper 1 must be connected to run this program.", "No connection", False, True, True)
                  end
                  if not(rq_is_gripper_activated("1")):
                    popup("Gripper 1 is not activated. Go to Installation tab > Gripper to activate it and run the program again.", "Not activated", False, True, True)
                  end
                  rq_set_pos_spd_for(255, 0, 77, "1")
                  rq_wait_pos_spe_for_request(255, 0, 77, "1")
                  rq_go_to("1")
                  rq_wait("1")
                  # end: URCap Program Node
                  $ 4480 "spat_flatS_up" "noBreak"
                  movel(spat_flatS_up_p, a=1.2, v=0.25, r=0.05)
                  $ 4481 "Spatula_otw" "noBreak"
                  movel(Spatula_otw_p, a=1.2, v=0.25)
                  $ 4482 "switch_spat_F_S≔ False " "noBreak"
                  global switch_spat_F_S=  False
                end
              end
            end
          end
        end
        $ 4483 "Action_Info≔'Scooping'" "noBreak"
        global Action_Info="Scooping"
        $ 4484 "auto_tilt_and_scoop(W_now, target_weight, weight_value)" "noBreak"
        auto_tilt_and_scoop(W_now, target_weight, weight_value)
        $ 4485 "Action_Info≔'Dosing'" "noBreak"
        global Action_Info="Dosing"
        # begin: URCap Program Node
        #   Source: SensoPart VISOR Robotic, 2.0.6, SensoPart Industriesensorik GmbH
        #   Type: Approach Pose
        $ 4486 "Approach Pose" "noBreak"
        movej(pose_trans(easyPickPose,p[0.0000,0.0000,-0.0000,0.0000,0.0000,0.0000]),a=0.2618,v=0.1745,t=0.000000,r=0.000000)
        # end: URCap Program Node
        # begin: URCap Program Node
        #   Source: SensoPart VISOR Robotic, 2.0.6, SensoPart Industriesensorik GmbH
        #   Type: Target Pose
        $ 4487 "Target Pose" "noBreak"
        movel(pose_trans(easyPickPose,p[0.0000,0.0000,-0.0000,0.0000,0.0000,0.0000]),a=0.0500,v=0.0200,t=0.000000,r=0.000000)
        # end: URCap Program Node
        $ 4488 "Close Gripper" "noBreak"
        $ 4489 "dispense_pos≔get_actual_tcp_pose()" "noBreak"
        global dispense_pos= get_actual_tcp_pose ()
        $ 4490 "Loop weight_value≤target_weight and delta_count<3" "noBreak"
        thread Thread_while_4490():
          while (True):
            $ 4491 "MoveL" "noBreak"
            $ 4492 "dispense_pos" "noBreak"
            movel(dispense_pos, a=0.2, v=0.1)
            $ 4493 "log_weight()" "noBreak"
            log_weight()
            $ 4494 "CCW_full_Rotate()" "noBreak"
            CCW_full_Rotate()
            $ 4495 "Wait: 0.5" "noBreak"
            sleep(0.5)
            $ 4496 "tilt_pose≔pose_trans(get_actual_tcp_pose(), p[0, 0, 0, 0, 0, 2.0])" "noBreak"
            global tilt_pose=pose_trans(get_actual_tcp_pose(), p[0, 0, 0, 0, 0, 2.0])
            $ 4497 "movel(tilt_pose, a=0.5, v=0.5, r=0.00001)" "noBreak"
            movel(tilt_pose, a=0.5, v=0.5, r=0.00001)
            $ 4498 "weight_value≔get_weight()" "noBreak"
            global weight_value=get_weight()
            $ 4499 "tilt_angle≔-1" "noBreak"
            global tilt_angle=-1
            $ 4500 "Wait: 0.5" "noBreak"
            sleep(0.5)
            $ 4501 "dispense_pos" "noBreak"
            movel(dispense_pos, a=1.2, v=0.25)
            $ 4502 "compute_level_percent(W_now, weight_value)" "noBreak"
            compute_level_percent(W_now, weight_value)
            $ 4503 "If delta<0.01" "noBreak"
            if (delta<0.01):
              $ 4504 "delta_count≔delta_count+1" "noBreak"
              global delta_count=delta_count+1
            else:
              $ 4505 "Else" "noBreak"
              $ 4506 "delta_count≔0" "noBreak"
              global delta_count=0
            end
            $ 4507 "prev_spat≔spatula" "noBreak"
            global prev_spat=spatula
            $ 4508 "Wait: 0.2" "noBreak"
            sleep(0.2)
            $ 4509 "spatula≔select_spatula(Flowability, level, diff, bulk_density, mouth_d)" "noBreak"
            global spatula=select_spatula(Flowability, level, diff, bulk_density, mouth_d)
            $ 4510 "Wait: 1.0" "noBreak"
            sleep(1.0)
            $ 4511 "send_level_info()" "noBreak"
            send_level_info()
            $ 4512 "send_spatula_info()" "noBreak"
            send_spatula_info()
            $ 4513 "Set AO[0]=0.0" "noBreak"
            set_standard_analog_out(0, 0.0)
            $ 4514 "Wait: 0.5" "noBreak"
            sleep(0.5)
            $ 4515 "swtich spatula" "noBreak"
            $ 4516 "If spatula ≟ 'spatula_M' and switch_spat_M≟ True " "noBreak"
            if (spatula  ==  "spatula_M"  and  switch_spat_M ==   True  ):
              $ 4517 "MoveJ" "noBreak"
              $ 4518 "Spatula_otw" "noBreak"
              movej(get_inverse_kin(Spatula_otw_p, qnear=Spatula_otw_q), a=1.3962634015954636, v=1.0471975511965976)
              $ 4519 "spat_L_up" "noBreak"
              movej(get_inverse_kin(spat_L_up_p, qnear=spat_L_up_q), a=1.3962634015954636, v=1.0471975511965976)
              $ 4520 "MoveL" "noBreak"
              $ 4521 "spat_L_side" "noBreak"
              movel(spat_L_side_p, a=1.2, v=0.25)
              $ 4522 "spat_L_lift" "noBreak"
              movel(spat_L_lift_p, a=1.2, v=0.25)
              $ 4523 "spat_L_pick" "noBreak"
              movel(spat_L_pick_p, a=0.2, v=0.1)
              # begin: URCap Program Node
              #   Source: Robotiq_Grippers, 3.17.0.105337, Robotiq Inc.
              #   Type: Gripper
              $ 4524 "Gripper Open (1)" "noBreak"
              if not(gripper_connected[0]):
                popup("Gripper 1 must be connected to run this program.", "No connection", False, True, True)
              end
              if not(rq_is_gripper_activated("1")):
                popup("Gripper 1 is not activated. Go to Installation tab > Gripper to activate it and run the program again.", "Not activated", False, True, True)
              end
              rq_set_pos_spd_for(0, 255, 77, "1")
              rq_wait_pos_spe_for_request(0, 255, 77, "1")
              rq_go_to("1")
              rq_wait("1")
              # end: URCap Program Node
              $ 4525 "spat_M_pick" "noBreak"
              movel(spat_M_pick_p, a=1.2, v=0.25)
              # begin: URCap Program Node
              #   Source: Robotiq_Grippers, 3.17.0.105337, Robotiq Inc.
              #   Type: Gripper
              $ 4526 "Gripper Close (1)" "noBreak"
              if not(gripper_connected[0]):
                popup("Gripper 1 must be connected to run this program.", "No connection", False, True, True)
              end
              if not(rq_is_gripper_activated("1")):
                popup("Gripper 1 is not activated. Go to Installation tab > Gripper to activate it and run the program again.", "Not activated", False, True, True)
              end
              rq_set_pos_spd_for(255, 0, 77, "1")
              rq_wait_pos_spe_for_request(255, 0, 77, "1")
              rq_go_to("1")
              rq_wait("1")
              # end: URCap Program Node
              $ 4527 "spat_M_up" "noBreak"
              movel(spat_M_up_p, a=1.2, v=0.25)
              $ 4528 "Spatula_otw" "noBreak"
              movel(Spatula_otw_p, a=1.2, v=0.25)
              $ 4529 "switch_spat_M≔ False " "noBreak"
              global switch_spat_M=  False
              $ 4530 "correction_reset()" "noBreak"
              correction_reset()
            else:
              $ 4531 "ElseIf spatula ≟ 'spatula_S' and switch_spat_S ≟ True and prev_spat≟'spatula_M'" "noBreak"
              if (spatula  ==  "spatula_S" and switch_spat_S  ==   True  and prev_spat == "spatula_M"):
                $ 4532 "MoveL" "noBreak"
                $ 4533 "Spatula_otw" "noBreak"
                movel(Spatula_otw_p, a=1.2, v=0.25)
                $ 4534 "spat_M_up" "noBreak"
                movel(spat_M_up_p, a=1.2, v=0.25)
                $ 4535 "spat_M_pick" "noBreak"
                movel(spat_M_pick_p, a=0.2, v=0.1)
                # begin: URCap Program Node
                #   Source: Robotiq_Grippers, 3.17.0.105337, Robotiq Inc.
                #   Type: Gripper
                $ 4536 "Gripper Open (1)" "noBreak"
                if not(gripper_connected[0]):
                  popup("Gripper 1 must be connected to run this program.", "No connection", False, True, True)
                end
                if not(rq_is_gripper_activated("1")):
                  popup("Gripper 1 is not activated. Go to Installation tab > Gripper to activate it and run the program again.", "Not activated", False, True, True)
                end
                rq_set_pos_spd_for(0, 255, 77, "1")
                rq_wait_pos_spe_for_request(0, 255, 77, "1")
                rq_go_to("1")
                rq_wait("1")
                # end: URCap Program Node
                $ 4537 "spat_S_pick" "noBreak"
                movel(spat_S_pick_p, a=1.2, v=0.25)
                # begin: URCap Program Node
                #   Source: Robotiq_Grippers, 3.17.0.105337, Robotiq Inc.
                #   Type: Gripper
                $ 4538 "Gripper Close (1)" "noBreak"
                if not(gripper_connected[0]):
                  popup("Gripper 1 must be connected to run this program.", "No connection", False, True, True)
                end
                if not(rq_is_gripper_activated("1")):
                  popup("Gripper 1 is not activated. Go to Installation tab > Gripper to activate it and run the program again.", "Not activated", False, True, True)
                end
                rq_set_pos_spd_for(255, 0, 77, "1")
                rq_wait_pos_spe_for_request(255, 0, 77, "1")
                rq_go_to("1")
                rq_wait("1")
                # end: URCap Program Node
                $ 4539 "spat_S_up" "noBreak"
                movel(spat_S_up_p, a=1.2, v=0.25)
                $ 4540 "Spatula_otw" "noBreak"
                movel(Spatula_otw_p, a=1.2, v=0.25)
                $ 4541 "switch_spat_S≔ False " "noBreak"
                global switch_spat_S=  False
                $ 4542 "correction_reset()" "noBreak"
                correction_reset()
              else:
                $ 4543 "ElseIf spatula≟'spatula_S' and switch_spat_S≟ True  and prev_spat≟'spatula_L'" "noBreak"
                if (spatula == "spatula_S" and switch_spat_S ==   True    and  prev_spat == "spatula_L"):
                  $ 4544 "MoveJ" "noBreak"
                  $ 4545 "Spatula_otw" "noBreak"
                  movej(get_inverse_kin(Spatula_otw_p, qnear=Spatula_otw_q), a=1.3962634015954636, v=1.0471975511965976)
                  $ 4546 "spat_L_up" "noBreak"
                  movej(get_inverse_kin(spat_L_up_p, qnear=spat_L_up_q), a=1.3962634015954636, v=1.0471975511965976)
                  $ 4547 "MoveL" "noBreak"
                  $ 4548 "spat_L_side" "noBreak"
                  movel(spat_L_side_p, a=1.2, v=0.25)
                  $ 4549 "spat_L_lift" "noBreak"
                  movel(spat_L_lift_p, a=1.2, v=0.25)
                  $ 4550 "spat_L_pick" "noBreak"
                  movel(spat_L_pick_p, a=0.2, v=0.1)
                  # begin: URCap Program Node
                  #   Source: Robotiq_Grippers, 3.17.0.105337, Robotiq Inc.
                  #   Type: Gripper
                  $ 4551 "Gripper Open (1)" "noBreak"
                  if not(gripper_connected[0]):
                    popup("Gripper 1 must be connected to run this program.", "No connection", False, True, True)
                  end
                  if not(rq_is_gripper_activated("1")):
                    popup("Gripper 1 is not activated. Go to Installation tab > Gripper to activate it and run the program again.", "Not activated", False, True, True)
                  end
                  rq_set_pos_spd_for(0, 255, 77, "1")
                  rq_wait_pos_spe_for_request(0, 255, 77, "1")
                  rq_go_to("1")
                  rq_wait("1")
                  # end: URCap Program Node
                  $ 4552 "spat_S_pick" "noBreak"
                  movel(spat_S_pick_p, a=1.2, v=0.25)
                  # begin: URCap Program Node
                  #   Source: Robotiq_Grippers, 3.17.0.105337, Robotiq Inc.
                  #   Type: Gripper
                  $ 4553 "Gripper Close (1)" "noBreak"
                  if not(gripper_connected[0]):
                    popup("Gripper 1 must be connected to run this program.", "No connection", False, True, True)
                  end
                  if not(rq_is_gripper_activated("1")):
                    popup("Gripper 1 is not activated. Go to Installation tab > Gripper to activate it and run the program again.", "Not activated", False, True, True)
                  end
                  rq_set_pos_spd_for(255, 0, 77, "1")
                  rq_wait_pos_spe_for_request(255, 0, 77, "1")
                  rq_go_to("1")
                  rq_wait("1")
                  # end: URCap Program Node
                  $ 4554 "spat_S_up" "noBreak"
                  movel(spat_S_up_p, a=1.2, v=0.25)
                  $ 4555 "Spatula_otw" "noBreak"
                  movel(Spatula_otw_p, a=1.2, v=0.25)
                  $ 4556 "switch_spat_S≔ False " "noBreak"
                  global switch_spat_S=  False
                  $ 4557 "correction_reset()" "noBreak"
                  correction_reset()
                else:
                  $ 4558 "ElseIf spatula≟'spatula_flat_S'  and switch_spat_F_S ≟ True " "noBreak"
                  if (spatula == "spatula_flat_S"   and  switch_spat_F_S  ==   True  ):
                    $ 4559 "MoveL" "noBreak"
                    $ 4560 "Spatula_otw" "noBreak"
                    movel(Spatula_otw_p, a=1.2, v=0.25)
                    $ 4561 "spat_flatM_up" "noBreak"
                    movel(spat_flatM_up_p, a=1.2, v=0.25)
                    $ 4562 "spat_flatM_pick" "noBreak"
